(* IEC 61131-3 sources: daoli-st-library/DL_Motion (part 14) *)

(* ---- FB_DL_GearDecouple.st ---- *)
(*==============================================================================
 * 组件名称 (Component)  : FB_DL_GearDecouple
 * 所属子库 (Sublibrary) : DL_Motion
 * 当前版本 (Version)    : 1.0.0
 * 兼容性   (Platform)   : CODESYS 3.5+ / TwinCAT 3 / 汇川 InoProShop / 施耐德 Machine Expert
 *                         仅依赖 Standard.library（ABS），零厂商私有库
 * 功能描述 (Function)   : 电子齿轮渐变脱耦（MC_GearOut 语义）：耦合期输出比例
 *                         fRatioOut = iNum ÷ iDen；脱耦请求（bCoupled 下降沿）
 *                         后比例按 tRamp 渐降至 1:1（禁直接跳断，规格指定），
 *                         到达 1:1 置 bReleased（电平指示，重耦合撤销）；脱耦
 *                         斜坡中重新耦合（bCoupled 上升沿）比例斜坡回升至全
 *                         比例，无阶跃。iDen = 0 → 拒绝并锁存故障（除数前置
 *                         闸，规格指定）。
 * 接口     (Interface)  : 输入 bCoupled 耦合命令（TRUE=全比例耦合）、iNum 齿轮
 *                         分子、iDen 齿轮分母（域 <> 0）、fRampS 脱耦渐变时长
 *                         （域 > 0） [s]、fCycle 扫描周期（<=0 用缺省） [s]、
 *                         bReset 复位；输出 fRatioOut 渐变比例、bReleased
 *                         脱耦完成指示（电平）、bRamping 斜坡执行中指示、
 *                         eErrCode 错误码、bError 故障标志。
 * 边界     (Boundary)   : ① **属主边界（写死）：本件只出渐变比例标量，不接管
 *                         轴使能、不下齿轮指令**；齿轮耦合执行归
 *                         `FB_DL_ElectronicGear`。
 *                         ② 斜率口径：全比例 fRatioFull = iNum/iDen，斜坡速率
 *                         = (fRatioFull − 1) ÷ fRampS [1/s]；单步 = 速率 × fCy，
 *                         步内可达即贴目标（无过冲）；fRampS 用 LREAL 秒口径，
 *                         避免跨平台 TIME→实数转换链（R64 交付门槛规避，头注释
 *                         声明工程取舍）。
 *                         ③ fRatioFull = 1（1:1 齿轮）时斜坡速率恒 0：脱耦
 *                         请求即达 1:1，当拍 bReleased（无跳变路径，比例本就
 *                         不变）。
 *                         ④ 斜坡中禁直接跳断：bCoupled 变化只改目标值，输出
 *                         恒限步逼近（头注释声明，规格指定）。
 *                         ⑤ 组态闸：iDen = 0 或 fRampS <= 0 → 锁存故障，输出
 *                         冻结保持末值（比例冻结语义声明：R191 二选一之「冻结
 *                         保持」，故障期禁跳变），解除沿 = bReset 上升沿。
 *                         ⑥ 非有限判据（R79 双判）：fCycle 非有限按缺省周期
 *                         处理并入组态闸（iNum/iDen 整型无浮点域）。
 *                         ⑦ 零全局耦合（无 GVL / VAR_EXTERNAL / 物理地址）。
 * 分工声明 (Scope)      : 与 `FB_DL_ElectronicGear` 分工：恒比例齿轮耦合归那件、
 *                         渐变脱耦编排归本件；与 `FB_DL_AxisSynchronizedStop`
 *                         分工：同步停止归那件。
 * 来源标签 (Source Tag) : T1-6 ◐（PLCopen MC 语义只借 GearOut 脱耦完成语义，
 *                         斜坡渐变实现为道莅自研 clean-room）
 * 码表     (Codes)      : 本件不占用任何全局数字码位。出口为 LREAL 比例 +
 *                         BOOL 组 + ENUM 错误码；数字码位待主控收口阶段统一
 *                         派号。
 * 红线自检 (Redline)    : R1 ✓ 零 GVL/VAR_EXTERNAL ｜ R2 ✓ 零 %I/%Q/%M ｜ R3 ✓ 纯 IEC 61131-3
 *                         R4 ✓ 除数前置闸 + 限步逼近 + 故障冻结声明 ｜ R5 ✓ 声明逐行同行双语注释
 *                         R6 N/A（锁存态无 CASE 状态机） ｜ R7 ✓ 一 R_TRIG 段 0 无条件刷新
 * 修订历史 (Revision)   : 2026-11-20  v1.0.0  R50 首版（批次 3 · 序号 14）
 * 验收向量 (Acceptance) : ① iNum=2, iDen=1（全比例 2.0），fRampS=2.0，
 *                         fCycle=0.01 → 单步 0.005：脱耦后 200 拍达 1.0 →
 *                         bReleased=TRUE；② 100 拍时重耦合 → 比例自 1.5 反向
 *                         斜坡回升至 2.0（无阶跃）；③ iDen=0 → 锁存 eCfgBad，
 *                         fRatioOut 冻结末值；④ iNum=1, iDen=1 → 脱耦请求
 *                         当拍 fRatioOut=1.0、bReleased=TRUE。
 *==============================================================================*)

(*-----------------------------------------------------------------------------
 * 枚举: E_DL_GdcErr（错误码；故障级恒伴 bError=TRUE）
 *----------------------------------------------------------------------------*)
TYPE E_DL_GdcErr :
(
    eOk     := 0,   // 正常 / Normal
    eCfgBad := 1    // 故障级：分母零或斜坡时长非法（输出冻结保持） / Fault: zero denominator or bad ramp time
);
END_TYPE

FUNCTION_BLOCK FB_DL_GearDecouple
VAR_INPUT
    bCoupled : BOOL := TRUE;          // 耦合命令（TRUE=全比例，FALSE=脱耦请求） [-] / Coupled command
    iNum     : DINT := 2;             // 齿轮分子 [-] / Gear numerator
    iDen     : DINT := 1;             // 齿轮分母，域 <> 0 [-] / Gear denominator, must not be zero
    fRampS   : LREAL := 2.0;          // 脱耦渐变时长（全比例→1:1），域 > 0 [s] / Decouple ramp duration [s]
    fCycle   : LREAL := 0.0;          // 扫描周期（<=0 用缺省） [s] / Scan cycle, default used when <= 0
    bReset   : BOOL := FALSE;         // 复位，上升沿清组态锁存并回全比例/1:1 目标重算 [-] / Reset, rising edge clears latch
END_VAR
VAR_OUTPUT
    fRatioOut : LREAL;                // 渐变比例输出（限步逼近目标） [-] / Ramped ratio output
    bReleased : BOOL;                 // 脱耦完成指示（比例达 1:1 ∧ 脱耦请求中，电平） [-] / Released indicator, level
    bRamping  : BOOL;                 // 斜坡执行中指示 [-] / Ramping indicator
    eErrCode  : E_DL_GdcErr;          // 错误码出口 / Error code outlet
    bError    : BOOL;                 // 故障标志（组态锁存） [-] / Error flag, latched
END_VAR
VAR
    _fRatio   : LREAL := 1.0;         // 比例内部锁存（限步源，初值 1:1 安全态） / Ratio internal latch
    _fFull    : LREAL;                // 全比例 = iNum ÷ iDen（分母已闸） [-] / Full ratio
    _fRate    : LREAL;                // 斜坡速率（全比例−1）÷fRampS [1/s] / Ramp rate
    _fStep    : LREAL;                // 当拍最大步长 [1/拍] / Max step this scan
    _fTarget  : LREAL;                // 当拍目标比例 [-] / Target ratio this scan
    _fCy      : LREAL;                // 当拍有效周期 [s] / Effective cycle this scan
    _bCfgBad  : BOOL;                 // 组态非法当拍量 [-] / Illegal configuration
    _bErrLatch: BOOL;                 // 组态故障锁存位（解除沿 = bReset 上升沿） / Latched config fault
    rtReset   : R_TRIG;               // 复位沿实例，段 0 无条件调用 / Reset edge instance
END_VAR
VAR CONSTANT
    DL_GDC_CYDEF : LREAL := 0.01;     // 缺省扫描周期 [s] / Default scan cycle
    DL_GDC_ONE   : LREAL := 1.0;      // 1:1 基准与到达容差中心 [-] / Unity ratio base
    DL_GDC_ZERO  : LREAL := 0.0;      // 判零基准 [-] / Zero base
    DL_GDC_TOL   : LREAL := 1.0E-6;   // 到达判据容差（浮点禁 = 判等） [-] / Arrival tolerance
END_VAR

(* —— 段 0：非有限判 + 组态闸 + 周期派生 + 沿刷新 —— *)
IF fCycle <> fCycle THEN
    _fCy := DL_GDC_CYDEF;                          // 周期非有限按缺省（规格⑥） / Non-finite cycle to default
ELSIF fCycle > DL_GDC_ZERO THEN
    _fCy := fCycle;                                // 组态周期有效 / Configured cycle
ELSE
    _fCy := DL_GDC_CYDEF;                          // 周期缺省兜底 / Default fallback
END_IF
_bCfgBad := (iDen = 0) OR (fRampS <= DL_GDC_ZERO);   // 组态域闸（除数前置 + 斜坡时长） / Configuration gate
rtReset(CLK := bReset);                            // 复位沿，每拍必调 / Reset edge, every scan

(* —— 段 1：复位沿与组态锁存 —— *)
IF rtReset.Q THEN
    _bErrLatch := FALSE;                           // 清组态锁存（R188 声明：解除沿 = bReset 上升沿） / Clear cfg latch
END_IF
IF _bCfgBad AND (NOT _bErrLatch) THEN
    _bErrLatch := TRUE;                            // 锁存 / Latch
END_IF

(* —— 段 2：目标与速率派生（故障期跳过派生，冻结保持） —— *)
IF NOT _bErrLatch THEN
    _fFull := DINT_TO_LREAL(iNum) / DINT_TO_LREAL(iDen);   // 全比例（分母已闸，无除零） / Full ratio
    _fRate := ABS(_fFull - DL_GDC_ONE) / fRampS;   // 斜坡速率（对称双向同一速率） / Ramp rate
    _fStep := _fRate * _fCy;                       // 单步上限 [1/拍] / Max step
    IF bCoupled THEN
        _fTarget := _fFull;                        // 耦合目标 = 全比例 / Coupled target
    ELSE
        _fTarget := DL_GDC_ONE;                    // 脱耦目标 = 1:1（MC_GearOut 语义） / Decouple target
    END_IF
END_IF

(* —— 段 3：限步逼近（斜坡中禁直接跳断，规格④；步内可达即贴目标） —— *)
IF NOT _bErrLatch THEN
    IF _fTarget > (_fRatio + _fStep) THEN
        _fRatio := _fRatio + _fStep;               // 正向限步（重耦合回升无阶跃） / Ramp up limited
    ELSIF _fTarget < (_fRatio - _fStep) THEN
        _fRatio := _fRatio - _fStep;               // 负向限步（脱耦渐降） / Ramp down limited
    ELSE
        _fRatio := _fTarget;                       // 步内到达：贴目标 / Settle at target
    END_IF
END_IF

(* —— 段 4：出口单点映射（名实双出口同源，R191） —— *)
fRatioOut := _fRatio;                              // 比例出口（故障期冻结保持末值，头注释⑤声明） / Ratio outlet, frozen on fault
IF (NOT _bErrLatch) AND (NOT bCoupled)
   AND (ABS(_fRatio - DL_GDC_ONE) < DL_GDC_TOL) THEN
    bReleased := TRUE;                             // 脱耦完成电平（比例达 1:1 ∧ 脱耦请求中） / Released level
ELSE
    bReleased := FALSE;                            // 未完成/重耦合/故障期撤销 / Not released
END_IF
bRamping := (NOT _bErrLatch)
        AND (ABS(_fRatio - _fTarget) >= DL_GDC_TOL);   // 斜坡执行中（与目标距离超容差） / Ramping indicator
IF _bErrLatch THEN
    bError := TRUE;                                // 故障标志（R45 配对） / Error flag
    eErrCode := E_DL_GdcErr.eCfgBad;               // 故障级码 / Fault code
ELSE
    bError := FALSE;                               // 无故障级条件 / No fault
    eErrCode := E_DL_GdcErr.eOk;                   // 正常码 / OK code
END_IF

END_FUNCTION_BLOCK

(* ---- FB_DL_GearHobAxialShiftSeq.st ---- *)
//==============================================================================
// 功能块：FB_DL_GearHobAxialShiftSeq ｜ 中文名称：滚齿机滚刀轴向窜刀顺控（复杂度 C4）
// 所属子库：DL_Motion ｜ 版本 VERSION: v1.0.0 ｜ 兼容：CODESYS V3.5+ / TwinCAT 3 / 汇川 InoProShop
// 功能描述：滚刀磨损后沿刀轴窜动一个切削区宽度换新切削区——松刀轴夹紧 → 轴向进给
//           到目标位 → 到位稳定 → 重新夹紧确认 → 对刀校验 → 完成，累计窜刀量在完成
//           拍提交；超可用行程拒动、未松夹不得进给、未夹紧不得对刀、步超时落故障；
//           中止走两段化（先停进给 → 轴静止窗 → 再按安全序重新夹紧）。
// 开源溯源 (Origin)：道莅原创实现（参考 GB/T 1356 圆柱齿轮滚齿工艺与滚刀轴向窜刀
//           量工程惯例 分类与参数域，许可证=MIT，借鉴点=「按切削区宽度分步窜刀并
//           累计至刀轴可用行程上限」的工艺序）
// 单位表：长度[mm] / 时间[ms] / 计数[次]
// 错误码表（Motion 段 0008，故障窗口 0A01~0A08，信息窗口 0101）：
//   16#0008_0A01 故障级：组态非法（步长/上限/容差 <= 0、累计初值 < 0、时间量 <= 0）
//   16#0008_0A02 故障级：目标位 > fMaxTravelMm，拒动并置 xTravelLimit
//   16#0008_0A03 故障级：松夹相超时未到位，或进给期松夹信号丢失，禁进给
//   16#0008_0A04 故障级：夹紧相或中止再夹紧窗超时未确认，禁对刀
//   16#0008_0A05 故障级：进给步超时，或稳定窗满仍未判轴到位
//   16#0008_0A06 故障级：轴位置入口非有限（NaN / Inf）或幅值超合法上限，拒算
//   16#0008_0A07 故障级：对刀校验偏差 > fPosTolMm
//   16#0008_0A08 故障级兜底：状态机落 ELSE 非法态，全输出断
//   16#0008_0101 信息级：单步窜刀完成（完成拍，不置 bError）
//           故障级码全部锁存回放（R187），唯一清除路径 = bReset 上升沿。
// 状态机：E_DL_HobShiftState（八态：eIdle=0 / eRelease=10 / eShift=20 / eSettle=30 /
//           eReclamp=40 / eVerify=50 / eDone=60 / eFault=99）。八态为纯相序机，中止
//           两段化不占相位（八态契约锁定），由内部段号 _uAbortStage 驱动（0 无 /
//           1 已停进给待轴静止 / 2 再夹紧中）。
// 边界行为：① 组态非法与入口非有限一律锁存故障，故障相不按当下输入重推断；② 故障
//           相迁出唯一路径 = bReset 上升沿且组态合法、未超程；③ 中止段 A 拍内
//           xCmdMove 立即断、夹紧两命令均不动（O 型中位液压锁保持），机检断言：中止
//           段 A 不得出现 xClampCmd / xUnclampCmd 置位；④ 八态 CASE 每态显式 + ELSE
//           兜底 → 0A08 全断；⑤ 目标位在启动拍锁定一次。
// 语义假设：① fTotalShiftMm 为累计窜刀量初值，只在首扫且未窜过刀时载入内部累计量，
//           运行期不参与运算（避免累计量双属主），掉电保持由上层把 fShiftUsedMm 回写
//           该引脚，且只允许在 eIdle 且 xStart = FALSE 期间回写；② 夹紧电磁阀为双电控
//           O 型中位机能——两命令全 FALSE 时液压锁保持，故故障相「全输出断」不会松开
//           刀轴；③ 位置反馈为刀轴轴向绝对位 [mm]，正方向为离开主轴端面的窜刀方向。
// 依赖纪律：仅 Standard.library（TON / R_TRIG）；零 GVL、零 VAR_EXTERNAL、零物理地
//           址直连，业务侧只经引脚注入。
// 修订历史：v1.0.0 2026-11-25 R88 首版（无人值守批次 · 复杂件 C4 · 序号 1）
//==============================================================================

(*------------------------------------------------------------------------------
 * 枚举: E_DL_HobShiftState（归属本功能块，同文件发布，全库唯一定义）
 * 含义: 窜刀顺控相位，与段 8 输出置位、段 9 码映射一一对应。
 *-----------------------------------------------------------------------------*)
TYPE E_DL_HobShiftState :
(
    eIdle    := 0,   // 空闲：等启动沿 / Idle, awaiting the start edge
    eRelease := 10,  // 松夹：发松开命令并等松开到位 / Release the arbor clamp and wait for feedback
    eShift   := 20,  // 轴向进给：发运动命令至目标位 / Axial feed towards the target position
    eSettle  := 30,  // 到位稳定：等稳定窗与到位标志 / Settle, stability window and in-position flag
    eReclamp := 40,  // 夹紧确认：发夹紧命令并等夹紧反馈 / Reclamp and wait for clamp feedback
    eVerify  := 50,  // 对刀校验：实测位与目标位比对 / Tool-position verification against the target
    eDone    := 60,  // 完成：累计窜刀量已提交 / Done, accumulated shift committed
    eFault   := 99   // 故障：组态/超程/联锁/超时/非法态 / Fault, configuration, travel, interlock, timeout or illegal state
);
END_TYPE

FUNCTION_BLOCK FB_DL_GearHobAxialShiftSeq
VAR_INPUT
    xEnable       : BOOL;   // 使能，FALSE 期间按中止处理 [—] / Enable, a drop is treated as an abort
    xStart        : BOOL;   // 启动请求，上升沿生效 [—] / Start request, rising edge effective
    xAbort        : BOOL;   // 中止请求，任意拍生效 [—] / Abort request, effective on any scan
    xReset        : BOOL;   // 故障复位，上升沿清全部锁存 [—] / Fault reset, rising edge clears all latches
    fShiftStepMm  : LREAL;  // 单步窜刀量 [mm]，须 > 0 / Per-step axial shift [mm], must be > 0
    fTotalShiftMm : LREAL;  // 累计窜刀量初值 [mm]，仅首扫载入 / Initial accumulated shift [mm], first scan only
    fAxisPosMm    : LREAL;  // 刀轴实际轴向位置 [mm] / Hob arbor actual axial position [mm]
    xAxisInPos    : BOOL;   // 轴到位标志 [—] / Axis in-position flag
    xClampClosed  : BOOL;   // 夹紧到位反馈 [—] / Clamp-closed feedback
    xClampOpen    : BOOL;   // 松开到位反馈 [—] / Clamp-open feedback
    tMoveTimeout  : TIME;   // 进给/校验步超时 [ms] / Feed and verification step timeout [ms]
    tSettleTime   : TIME;   // 到位稳定窗 [ms] / In-position settle window [ms]
    fPosTolMm     : LREAL;  // 对刀位置容差 [mm]，须 > 0 / Verification position tolerance [mm]
    fMaxTravelMm  : LREAL;  // 刀轴可用窜刀总行程 [mm] / Total usable axial shift travel [mm]
END_VAR
VAR_OUTPUT
    xCmdMove      : BOOL;   // 轴向进给命令 [—] / Axial feed command
    fCmdPosMm     : LREAL;  // 目标位命令 [mm] / Target position command [mm]
    xClampCmd     : BOOL;   // 夹紧命令（双电控 O 型中位，断电保持） [—] / Clamp command, O-centre holds on power loss
    xUnclampCmd   : BOOL;   // 松开命令（双电控 O 型中位，断电保持） [—] / Unclamp command, holds on power loss
    bRunning      : BOOL;   // 顺控运行中（非空闲非完成非故障非中止） [—] / Sequencing active
    bDone         : BOOL;   // 单步窜刀完成相电平 [—] / Single shift step done, level in the done phase
    bError        : BOOL;   // 故障级标志，仅故障级码置位 [—] / Fault-class flag, fault-level codes only
    nErrCode      : UDINT;  // 错误码，0 = 无错 [—] / Error code, 0 = none
    fShiftUsedMm  : LREAL;  // 累计窜刀量出口 [mm] / Accumulated axial shift outlet [mm]
    nShiftCount   : UDINT;  // 累计窜刀次数 [次] / Accumulated shift step count
    xTravelLimit  : BOOL;   // 窜刀行程上限已达（拒动锁存） [—] / Travel limit reached, refuse-to-move latch
END_VAR
VAR
    _eState       : E_DL_HobShiftState := E_DL_HobShiftState.eIdle; // 当前相位 [—] / Current phase
    _bInit        : BOOL := FALSE;      // 首扫标志，取非判定 [—] / First-scan flag, tested negated
    _fShiftUsedMm : LREAL;              // 内部累计窜刀量 [mm] / Internal accumulated shift [mm]
    _fTargetPosMm : LREAL;              // 本步目标位 [mm] = 累计 + 步长 / Step target [mm] = accumulated + step
    _fPosPrevMm   : LREAL;              // 上拍轴位快照 [mm]，静止判据用 / Previous-scan position [mm]
    _nShiftCount  : UDINT;              // 内部累计窜刀次数 [次] / Internal shift step counter
    _bCfgBad      : BOOL;               // 组态非法锁存 / Illegal configuration latch
    _bCfgOk       : BOOL;               // 本拍组态合法（派生量不锁存） [—] / Configuration legal this scan, derived
    _bAxisBad     : BOOL;               // 轴位置非有限锁存 / Non-finite axis position latch
    _bOverTravel  : BOOL;               // 超窜刀行程锁存 / Over-travel latch
    _bReleaseTmo  : BOOL;               // 松夹未到位/信号丢失锁存 / Release-not-reached latch
    _bClampTmo    : BOOL;               // 夹紧未确认锁存 / Clamp-not-confirmed latch
    _bFeedTmo     : BOOL;               // 进给步超时锁存 / Feed step timeout latch
    _bVerifyErr   : BOOL;               // 对刀超差锁存 / Verification error latch
    _bIllegal     : BOOL;               // 非法状态标志 / Illegal state flag
    _bInfoDone    : BOOL;               // 单步完成信息当拍标志 / Step-done info flag of this scan
    _bAbortReq    : BOOL;               // 中止请求合成（xAbort 或失能） [—] / Combined abort request
    _bFeedPermit  : BOOL;               // 进给许可（松开到位且未夹紧） [—] / Feed permit, released and not clamped
    _bStandstill  : BOOL;               // 轴静止判据（本拍位移小于阈值） [—] / Axis standstill criterion
    _uAbortStage  : UINT;               // 中止段号 0=无 1=待静止 2=再夹紧 / Abort stage 0 none 1 standstill 2 reclamp
    rtStart       : R_TRIG;             // 启动沿，段 5 无条件刷新 [—] / Start edge, refreshed in segment 5
    rtReset       : R_TRIG;             // 复位沿，段 5 无条件刷新 [—] / Reset edge, refreshed in segment 5
    tonRelease    : TON;                // 松夹相超时计时 [ms] / Release phase timeout [ms]
    tonMove       : TON;                // 进给相超时计时 [ms] / Feed phase timeout [ms]
    tonSettle     : TON;                // 稳定窗计时 [ms] / Settle window timer [ms]
    tonReclamp    : TON;                // 夹紧确认超时计时 [ms] / Reclamp timeout [ms]
    tonVerify     : TON;                // 对刀校验超时计时 [ms] / Verification timeout [ms]
    tonStandstill : TON;                // 中止段 A 静止窗计时 [ms] / Abort stage A standstill window [ms]
    tonAbortClamp : TON;                // 中止段 B 再夹紧确认窗计时 [ms] / Abort stage B reclamp window [ms]
END_VAR
VAR CONSTANT
    DL_EPS           : LREAL := 1.0E-9;      // 浮点容差零点，兼作除法分母下限 / Float epsilon, also the divisor floor
    DL_HOB_STILL_MM  : LREAL := 0.005;       // 静止窗每拍位移阈值 [mm] / Per-scan displacement threshold [mm]
    DL_HOB_ABORT_T   : TIME  := T#1500MS;    // 中止静止窗时长 [ms] / Abort standstill window [ms]
    DL_HOB_CLAMP_T   : TIME  := T#3000MS;    // 中止再夹紧确认窗 [ms] / Abort reclamp confirm window [ms]
    DL_HOB_POS_MAX   : LREAL := 1.0E9;       // 位置幅值合法上限 [mm] / Legal position magnitude ceiling [mm]
END_VAR

(*------------------------------------------------------------------------------
 * 段 1｜每拍预置：全部输出先落安全侧，单拍标志预清零
 *      All outputs preset to the safe side, one-shot flags pre-cleared
 *-----------------------------------------------------------------------------*)
xCmdMove := FALSE;  fCmdPosMm := 0.0;       // 进给命令与目标位先清 / Feed command and target cleared first
xClampCmd := FALSE; xUnclampCmd := FALSE;   // 夹紧两命令先断（O 型中位保持） / Both clamp commands cleared, O-centre holds
bRunning := FALSE;  bDone := FALSE;         // 运行与完成标志每拍重算 / Running and done flags recomputed
bError := FALSE;    nErrCode := 16#0000_0000; // 故障标志与错误码每拍重算 / Fault flag and code recomputed
xTravelLimit := FALSE;                      // 超程标志每拍重算 / Travel limit flag recomputed
_bIllegal := FALSE; _bInfoDone := FALSE;    // 非法态与完成信息预清零 / Illegal and done-info flags pre-cleared

(*------------------------------------------------------------------------------
 * 段 2｜首扫初始化：相位、累计量、计数与中止段号复位
 *      First-scan initialisation of phase, accumulated shift, counter and abort stage
 *-----------------------------------------------------------------------------*)
IF NOT _bInit THEN
    _eState       := E_DL_HobShiftState.eIdle;   // 相位从空闲起步 / Phase starts idle
    _fShiftUsedMm := 0.0;  _fTargetPosMm := 0.0; // 累计量与目标位先清零 / Accumulated shift and target at zero
    _fPosPrevMm   := 0.0;  _nShiftCount  := 0;   // 位置快照与窜刀计数清零 / Position snapshot and counter at zero
    _uAbortStage  := 0;                          // 中止段号从零起步 / Abort stage starts at zero
    _bInit        := TRUE;                       // 首扫只做一次 / The first scan runs once
END_IF

(*------------------------------------------------------------------------------
 * 段 3｜入口非有限闸 + 组态闸 + 目标位预计算 + 超行程拒动判定
 *      Non-finite inlet gate, configuration gates, target computation, travel check
 *-----------------------------------------------------------------------------*)
IF NOT (fAxisPosMm > -1.0E30 AND fAxisPosMm < 1.0E30) THEN _bAxisBad := TRUE; END_IF    // 轴位非有限 → 0A06 / Non-finite position, 0A06
IF ABS(fAxisPosMm) > DL_HOB_POS_MAX THEN _bAxisBad := TRUE; END_IF                     // 轴位幅值超上限 → 0A06 / Beyond the ceiling, 0A06
IF NOT (fShiftStepMm > -1.0E30 AND fShiftStepMm < 1.0E30) THEN _bCfgBad := TRUE; END_IF  // 步长非有限 → 0A01 / Non-finite step, 0A01
IF NOT (fMaxTravelMm > -1.0E30 AND fMaxTravelMm < 1.0E30) THEN _bCfgBad := TRUE; END_IF // 行程上限非有限 → 0A01 / Non-finite limit, 0A01
IF NOT (fPosTolMm > -1.0E30 AND fPosTolMm < 1.0E30) THEN _bCfgBad := TRUE; END_IF      // 容差非有限 → 0A01 / Non-finite tolerance, 0A01
IF NOT (fTotalShiftMm > -1.0E30 AND fTotalShiftMm < 1.0E30) THEN _bCfgBad := TRUE; END_IF // 累计初值非有限 → 0A01 / Non-finite initial shift, 0A01
IF (fShiftStepMm <= DL_EPS) OR (fMaxTravelMm <= DL_EPS) OR (fPosTolMm <= DL_EPS) THEN _bCfgBad := TRUE; END_IF // 三者须为正 → 0A01 / All three must be positive
IF fTotalShiftMm < 0.0 THEN _bCfgBad := TRUE; END_IF                                   // 累计初值负值非法 → 0A01 / Negative initial shift, 0A01
IF (tMoveTimeout <= T#0MS) OR (tSettleTime <= T#0MS) THEN _bCfgBad := TRUE; END_IF      // 时间量须为正 → 0A01 / Time values must be positive
_bCfgOk := NOT _bCfgBad;                    // 本拍组态合法派生量 / Configuration-legal derived flag of this scan
IF (_nShiftCount = 0) AND (_eState = E_DL_HobShiftState.eIdle) AND (NOT _bCfgBad) THEN
    _fShiftUsedMm := fTotalShiftMm;         // 累计初值载入（仅未窜过刀时） / Initial shift loaded before the first step
END_IF
IF (_eState = E_DL_HobShiftState.eIdle) OR (_eState = E_DL_HobShiftState.eDone)
   OR (_eState = E_DL_HobShiftState.eFault) THEN
    _fTargetPosMm := _fShiftUsedMm + fShiftStepMm; // 目标位 = 累计窜刀量 + 步长 [mm]，仅非运行相更新，运行期锁定 / Target updated outside running phases only
END_IF
IF (_bCfgOk) AND (NOT _bAxisBad) AND (_fTargetPosMm > fMaxTravelMm) THEN
    _bOverTravel := TRUE;                   // 目标位超可利用行程，拒动锁存 → 0A02 / Beyond usable travel, 0A02
END_IF

(*------------------------------------------------------------------------------
 * 段 4｜中止入口（段 0→1）、静止判据与复位
 *      Abort entry, standstill criterion and the reset edge
 *-----------------------------------------------------------------------------*)
_bAbortReq   := xAbort OR (NOT xEnable);    // 中止请求合成：显式中止或失能 / Combined abort: explicit abort or enable loss
_bFeedPermit := xClampOpen AND (NOT xClampClosed); // 进给许可：松开到位且未夹紧 / Feed permit: released and not clamped
IF _bAbortReq AND (_uAbortStage = 0) AND (_eState <> E_DL_HobShiftState.eIdle)
   AND (_eState <> E_DL_HobShiftState.eDone) AND (_eState <> E_DL_HobShiftState.eFault) THEN
    _uAbortStage := 1;                      // 进中止段 A：先停进给待轴静止 / Enter abort stage A, await standstill
END_IF
_bStandstill := ABS(fAxisPosMm - _fPosPrevMm) < DL_HOB_STILL_MM; // 本拍位移小于阈值视为静止 / A per-scan move below the threshold is standstill
IF rtReset.Q THEN
    _bCfgBad := FALSE;  _bAxisBad := FALSE; _bOverTravel := FALSE; // 复位清组态/非有限/超程锁存 / Clears configuration, non-finite and travel
    _bReleaseTmo := FALSE; _bClampTmo := FALSE; _bFeedTmo := FALSE; // 复位清松夹/夹紧/超时锁存 / Clears release, clamp and timeout
    _bVerifyErr := FALSE;                   // 复位清对刀校验锁存 / Clears the verification latch
END_IF

(*------------------------------------------------------------------------------
 * 段 5｜定时器与边沿无条件周期刷新（R7：CASE 之外每拍必调，各司其职不复用）
 *      Timers and edges refreshed unconditionally every scan, outside the CASE
 *-----------------------------------------------------------------------------*)
rtStart(CLK := xStart);                     // 启动沿刷新 / Start edge refreshed
rtReset(CLK := xReset);                     // 复位沿刷新 / Reset edge refreshed
tonRelease(IN := (_eState = E_DL_HobShiftState.eRelease) AND (_uAbortStage = 0), PT := tMoveTimeout); // 松夹相超时 / Release timeout
tonMove(IN := (_eState = E_DL_HobShiftState.eShift) AND (_uAbortStage = 0), PT := tMoveTimeout);      // 进给相超时 / Feed timeout
tonSettle(IN := (_eState = E_DL_HobShiftState.eSettle) AND (_uAbortStage = 0), PT := tSettleTime);    // 稳定窗计时 / Settle window
tonReclamp(IN := (_eState = E_DL_HobShiftState.eReclamp) AND (_uAbortStage = 0), PT := tMoveTimeout); // 夹紧确认超时 / Reclamp timeout
tonVerify(IN := (_eState = E_DL_HobShiftState.eVerify) AND (_uAbortStage = 0), PT := tMoveTimeout);   // 对刀校验超时 / Verification timeout
tonStandstill(IN := (_uAbortStage = 1) AND _bStandstill, PT := DL_HOB_ABORT_T); // 中止段 A 静止窗 / Abort stage A standstill window
tonAbortClamp(IN := (_uAbortStage = 2), PT := DL_HOB_CLAMP_T);                  // 中止段 B 再夹紧窗 / Abort stage B reclamp window

(*------------------------------------------------------------------------------
 * 段 6｜中止段推进（1→2 轴静止后按安全序再夹紧，2→0 收口）
 *      Abort stage progression, reclamp only after the axis is standstill
 *-----------------------------------------------------------------------------*)
IF (_uAbortStage = 1) AND tonStandstill.Q THEN
    _uAbortStage := 2;                      // 轴静止窗满，进再夹紧段 / Standstill elapsed, enter reclamp
END_IF
IF _uAbortStage = 2 THEN
    IF xClampClosed THEN
        _uAbortStage := 0;                  // 再夹紧已确认，中止收口 / Reclamp confirmed, abort closed
        _eState      := E_DL_HobShiftState.eIdle; // 回空闲 / Back to idle
    ELSIF tonAbortClamp.Q THEN
        _bClampTmo   := TRUE;               // 再夹紧窗满无反馈 → 0A04 / Window elapsed without feedback, 0A04
        _uAbortStage := 0;                  // 中止段收口 / Abort stage closed
        _eState      := E_DL_HobShiftState.eFault; // 落故障 / Fall to fault
    END_IF
END_IF

(*------------------------------------------------------------------------------
 * 段 7｜状态机（中止期间迁移冻结；本段只做迁移，输出在段 8）
 *      Phase machine, transitions frozen while aborting, outputs in segment 8
 *-----------------------------------------------------------------------------*)
IF _uAbortStage = 0 THEN
    CASE _eState OF
        E_DL_HobShiftState.eIdle:           // 空闲：启动沿 + 组态合法 + 未超程才进松夹 / Idle, legal start edge only
            IF rtStart.Q AND _bCfgOk AND (NOT _bAxisBad) AND (NOT _bOverTravel) AND (NOT _bAbortReq) THEN
                _fTargetPosMm := _fShiftUsedMm + fShiftStepMm; // 启动拍锁定目标位 / Target locked at the start edge
                _eState := E_DL_HobShiftState.eRelease;        // 进松夹相 / To the release phase
            END_IF
        E_DL_HobShiftState.eRelease:        // 松夹：松开到位才允许进给 / Release, feeding only once released
            IF _bFeedPermit THEN _eState := E_DL_HobShiftState.eShift; // 松开到位，进进给相 / Released, to feed
            ELSIF tonRelease.Q THEN _bReleaseTmo := TRUE; _eState := E_DL_HobShiftState.eFault; // 超时未到位 → 0A03 / Timeout, 0A03
            END_IF
        E_DL_HobShiftState.eShift:          // 进给：松夹信号丢失即故障，到位进稳定相 / Feed, permit loss faults
            IF NOT _bFeedPermit THEN _bReleaseTmo := TRUE; _eState := E_DL_HobShiftState.eFault; // 松夹丢失 → 0A03 / Permit lost, 0A03
            ELSIF xAxisInPos THEN _eState := E_DL_HobShiftState.eSettle; // 到位，进稳定相 / In position, to settle
            ELSIF tonMove.Q THEN _bFeedTmo := TRUE; _eState := E_DL_HobShiftState.eFault; // 进给步超时 → 0A05 / Feed timeout, 0A05
            END_IF
        E_DL_HobShiftState.eSettle:         // 稳定：稳定窗满且仍到位才进夹紧 / Settle, reclamp after the window
            IF tonSettle.Q AND xAxisInPos THEN _eState := E_DL_HobShiftState.eReclamp; // 稳定到位，进夹紧 / Stable, to reclamp
            ELSIF tonSettle.Q THEN _bFeedTmo := TRUE; _eState := E_DL_HobShiftState.eFault; // 窗满未到位 → 0A05 / Elapsed, 0A05
            END_IF
        E_DL_HobShiftState.eReclamp:        // 夹紧：夹紧确认才允许对刀校验 / Reclamp, verification only once clamped
            IF xClampClosed AND (NOT xClampOpen) THEN _eState := E_DL_HobShiftState.eVerify; // 夹紧确认，进校验 / Clamped, verify
            ELSIF tonReclamp.Q THEN _bClampTmo := TRUE; _eState := E_DL_HobShiftState.eFault; // 超时未夹紧 → 0A04 / Clamp timeout, 0A04
            END_IF
        E_DL_HobShiftState.eVerify:         // 对刀校验：夹紧须保持，偏差在容差内即完成 / Verify with the clamp held
            IF NOT xClampClosed THEN _bClampTmo := TRUE; _eState := E_DL_HobShiftState.eFault; // 夹紧丢失 → 0A04 / Clamp lost, 0A04
            ELSIF ABS(fAxisPosMm - _fTargetPosMm) <= fPosTolMm THEN
                _fShiftUsedMm := _fShiftUsedMm + fShiftStepMm; // 完成拍提交累计窜刀量 / Accumulated shift committed
                _nShiftCount := _nShiftCount + 1; _bInfoDone := TRUE; // 次数递增 + 完成信息 / Counter plus done info
                _eState := E_DL_HobShiftState.eDone;           // 进完成相 / To the done phase
            ELSIF tonVerify.Q THEN _bVerifyErr := TRUE; _eState := E_DL_HobShiftState.eFault; // 超差 → 0A07 / Deviation, 0A07
            END_IF
        E_DL_HobShiftState.eDone:           // 完成：启动撤销且无中止请求才回空闲 / Done, back to idle once start drops
            IF (NOT xStart) AND (NOT _bAbortReq) THEN _eState := E_DL_HobShiftState.eIdle; END_IF
        E_DL_HobShiftState.eFault:          // 故障：复位沿且组态合法且未超程才回空闲 / Fault, reset edge only
            IF rtReset.Q AND _bCfgOk AND (NOT _bAxisBad) AND (NOT _bOverTravel) THEN _eState := E_DL_HobShiftState.eIdle; END_IF
        ELSE                                // 非法状态兜底（R6：CASE 必带 ELSE）/ Illegal-state fallback
            _bIllegal := TRUE; _eState := E_DL_HobShiftState.eFault; // 非法态 → 0A08，落故障 / Illegal state, 0A08
    END_CASE
END_IF

(*------------------------------------------------------------------------------
 * 段 8｜输出置位（次序即安全：进给受许可闸，夹紧两命令互斥）
 *      Output assignment, feed gated by the permit, clamp commands exclusive
 *-----------------------------------------------------------------------------*)
CASE _eState OF
    E_DL_HobShiftState.eRelease:            // 松夹相：只发松开命令 / Release phase, unclamp only
        xUnclampCmd := TRUE;                // 松开命令 / Unclamp command
    E_DL_HobShiftState.eShift:              // 进给相：命令位 + 进给许可双重闸 / Feed phase, target plus permit
        fCmdPosMm := _fTargetPosMm;         // 目标位命令 / Target position command
        xCmdMove  := _bFeedPermit;          // 未松夹到位不得进给 / Feeding forbidden unless released
    E_DL_HobShiftState.eSettle:             // 稳定相：保持命令位不撤 / Settle phase, command held
        fCmdPosMm := _fTargetPosMm;         // 目标位保持 / Target position held
    E_DL_HobShiftState.eReclamp:            // 夹紧相：只发夹紧命令 / Reclamp phase, clamp only
        xClampCmd := TRUE;                  // 夹紧命令 / Clamp command
    E_DL_HobShiftState.eDone:               // 完成相：完成电平 / Done phase, done level
        bDone := TRUE;                      // 单步完成 / Single step done
    ELSE                                    // 其余相（空闲/校验/故障）全断 / Other phases, all off
        xCmdMove := FALSE; xClampCmd := FALSE; xUnclampCmd := FALSE; // 全输出断 / All outputs off
END_CASE
IF _uAbortStage >= 1 THEN
    xCmdMove    := FALSE;                   // 中止段 A：进给立即断（安全侧） / Abort A, feed cut immediately
    xClampCmd   := FALSE; xUnclampCmd := FALSE; // 静止窗内两夹紧命令均不动（O 型中位保持） / Both idle in the window
    fCmdPosMm   := _fTargetPosMm;           // 命令位保持，禁回零溜刀 / Command held, no return-to-zero creep
    IF _uAbortStage = 2 THEN
        xClampCmd := NOT xClampClosed;      // 中止段 B：未夹紧则发夹紧（安全序） / Abort B, clamp unless clamped
    END_IF
END_IF
bRunning := (_eState <> E_DL_HobShiftState.eIdle) AND (_eState <> E_DL_HobShiftState.eDone)
            AND (_eState <> E_DL_HobShiftState.eFault) AND (_uAbortStage = 0); // 运行标志 / Running flag

(*------------------------------------------------------------------------------
 * 段 9｜出口量与错误码映射（锁存回放，R187：故障相不按当下输入重推断）
 *      Outlet quantities and the error-code map, latched replay
 *-----------------------------------------------------------------------------*)
fShiftUsedMm := _fShiftUsedMm;              // 累计窜刀量出口 [mm] / Accumulated shift outlet [mm]
nShiftCount  := _nShiftCount;               // 窜刀次数出口 [次] / Shift count outlet
xTravelLimit := _bOverTravel;               // 超程拒动出口 / Travel-limit outlet
IF _bIllegal THEN nErrCode := 16#0008_0A08; bError := TRUE;        // 故障级兜底：非法态 / Fault, illegal state fallback
ELSIF _bCfgBad THEN nErrCode := 16#0008_0A01; bError := TRUE;      // 故障级：组态非法 / Fault, illegal configuration
ELSIF _bAxisBad THEN nErrCode := 16#0008_0A06; bError := TRUE;     // 故障级：轴位非有限 / Fault, non-finite position
ELSIF _bOverTravel THEN nErrCode := 16#0008_0A02; bError := TRUE;  // 故障级：超窜刀行程 / Fault, over travel
ELSIF _bReleaseTmo THEN nErrCode := 16#0008_0A03; bError := TRUE;  // 故障级：松夹不到位 / Fault, release not reached
ELSIF _bClampTmo THEN nErrCode := 16#0008_0A04; bError := TRUE;    // 故障级：夹紧未确认 / Fault, clamp not confirmed
ELSIF _bFeedTmo THEN nErrCode := 16#0008_0A05; bError := TRUE;     // 故障级：进给步超时 / Fault, feed step timeout
ELSIF _bVerifyErr THEN nErrCode := 16#0008_0A07; bError := TRUE;   // 故障级：对刀超差 / Fault, verification out of tolerance
ELSIF _bInfoDone THEN nErrCode := 16#0008_0101;                    // 信息级：单步完成，不置 bError / Info, step done
END_IF
_fPosPrevMm := fAxisPosMm;                  // 位置快照推进（供下拍静止判据） / Position snapshot advanced for the next scan
END_FUNCTION_BLOCK

(* ---- FB_DL_GearInPhaseAlign.st ---- *)
(*
  FB_DL_GearInPhaseAlign  —  电子齿轮啮合相位对齐（相位差窗 + 从轴偏置补偿） / Electronic gear-in phase alignment with phase-error window and slave offset compensation
  分类 Category : DL_Motion
  版本 Version  : 1.0.0
  来源 Source   : t1-6-plcopen — PLCopen Motion 接口映射层族深化
  溯源 Origin   : 道莅 clean-room 实现；从轴相位 = 主轴位置×传动比 + 偏置 为公开电子齿轮运动学关系，
                 本件仅做 MC_GearIn 前置相位判据与偏置补偿的映射层，不内联轨迹规划内核
  功能 Function : 1) 理想从轴相位 _fIdealDeg = fMasterPosDeg × fGearRatio；
                  2) 相位差 _fPhaseErrDeg = 归一化(fSlavePosDeg - _fIdealDeg - fPhaseTargetDeg)，
                  归一化按 ±360° 折算（除以常量 360.0，禁 MOD 非标准扩展）；
                  3) 判据：|相位差| <= fPhaseTolDeg → bInPhase（可啮合）；
                  4) 偏置补偿：补偿量按 -相位差 × fGainDegPerDeg 计算，钳制到
                  ±fOffsetMaxDeg 并限速（单次不超过 fOffsetStepDeg）；
                  5) 本件只有故障码、无信息码（派单硬约束）。
  接口 Interface: 输入主轴/从轴位置、传动比、目标相位、容差、偏置域；输出相位差与偏置
  边界 Boundary : ① 组态闸：fGearRatio <= 0.0、fPhaseTolDeg <= 0.0、fOffsetMaxDeg <= 0.0、
                  fOffsetStepDeg <= 0.0、fGainDegPerDeg <= 0.0 → 04A7 锁存；
                  ② 位置或传动比非有限（NaN 自反 + Inf 差值自减）→ 04A7 锁存，偏置冻结保持；
                  ③ 归一化除法除数为常量 360.0（无除零风险）；
                  ④ 一个 R_TRIG，段 0 无条件调用；⑤ 故障相迁出唯一路径 = bReset 上升沿；
                  ⑥ 零全局耦合：无 GVL / VAR_EXTERNAL / %I %Q %M 直接地址。
  依赖 Depends  : Standard.library（R_TRIG）
  码表 Error codes（Motion 段 0004，故障窗口 04A7；本件无信息码）:
    16#0004_04A7 故障级：相位对齐故障总码（组态非法 / 位置或传动比非有限），
                 锁存至 bReset 上升沿；归因见 eCause，不新增码位（派单硬约束单码）
  修订历史 Revision :
    2026-11-19  v1.0.0  R43 首版（批次 4 · 序号 19）
*)

TYPE E_DL_GpaState :
(
    eIdle   := 0,     // 未使能待对齐 / Idle, waiting alignment
    eAlign  := 10,    // 相位对齐中（偏置补偿） / Aligning with offset compensation
    eReady  := 20,    // 相位在窗：可啮合 / In phase, gear-in permitted
    eFault  := 90     // 故障锁存相（偏置冻结） / Fault latched, offset frozen
);
END_TYPE

TYPE E_DL_GpaCause :
(
    eNone       := 0, // 无故障成因 / No cause
    eCfgIllegal := 1, // 组态非法 / Illegal configuration
    eNonFinite  := 2  // 输入非有限 / Non-finite input
);
END_TYPE

FUNCTION_BLOCK FB_DL_GearInPhaseAlign
VAR_INPUT
    fMasterPosDeg  : REAL := 0.0;      // 主轴位置 [°] / Master position
    fSlavePosDeg   : REAL := 0.0;      // 从轴位置 [°] / Slave position
    fGearRatio     : REAL := 1.0;      // 传动比 [从轴°/主轴°]，域 > 0 / Gear ratio
    fPhaseTargetDeg: REAL := 0.0;      // 目标相位差 [°] / Target phase difference
    fPhaseTolDeg   : REAL := 2.0;      // 相位差窗 [°]，域 > 0 / Phase window
    fGainDegPerDeg : REAL := 0.8;      // 补偿增益 [°/°]，域 > 0 / Compensation gain
    fOffsetMaxDeg  : REAL := 30.0;     // 偏置限幅 [°]，域 > 0 / Offset limit
    fOffsetStepDeg : REAL := 5.0;      // 单周期偏置步长 [°]，域 > 0 / Offset step
    bEnable        : BOOL := FALSE;    // 对齐使能（电平）[-] / Alignment enable
    bReset         : BOOL := FALSE;    // 复位命令，上升沿清故障与偏置 [-] / Reset edge
END_VAR
VAR_OUTPUT
    eState         : E_DL_GpaState;    // 状态出口，段 6 单点映射 / State outlet
    eCause         : E_DL_GpaCause;    // 故障成因出口（R190） / Fault cause outlet
    fPhaseErrDeg   : REAL;             // 归一化相位差 [°] / Normalised phase error
    fOffsetDeg     : REAL;             // 从轴偏置补偿 [°] / Slave offset compensation
    bInPhase       : BOOL;             // 相位在窗（MC_GearIn 许可）[-] / In-phase permit
    bError         : BOOL;             // 故障锁存标志 [-] / Fault latch flag
    nErrId         : UDINT;            // 故障码，0 = 无故障（本件无信息码） / Fault code only
END_VAR
VAR
    _eState        : E_DL_GpaState := E_DL_GpaState.eIdle;   // 内部相位（CASE 唯一写入目标） / Internal phase
    _eCause        : E_DL_GpaCause := E_DL_GpaCause.eNone;   // 故障成因锁存（锁存量） / Latched cause
    rtReset        : R_TRIG;           // 复位沿实例，每周期无条件调用 / Reset edge
    _fOffsetDeg    : REAL;             // 偏置保持量（持久） / Offset holding slot
    _fIdealDeg     : REAL;             // 理想从轴相位 [°]（当拍量） / Ideal slave phase
    _fErrRawDeg    : REAL;             // 未归一化相位差 [°]（当拍量） / Raw phase error
    _fErrDeg       : REAL;             // 归一化相位差 [°]（当拍量） / Normalised phase error
    _fCmdDeg       : REAL;             // 目标偏置 [°]（当拍量） / Target offset
    _bInPhase      : BOOL;             // 相位在窗当拍量 [-] / In-phase verdict
    _bNonFin       : BOOL;             // 输入非有限当拍量 [-] / Non-finite input
    _bCfgBad       : BOOL;             // 组态非法当拍量 [-] / Config illegal
    _bFault        : BOOL;             // 故障锁存位（锁存量） / Latched fault bit
    _uFault        : UDINT;            // 故障码锁存（锁存量） / Latched fault code
END_VAR

(* —— 段 0：沿实例无条件周期刷新 + 相位差归一化（除数为常量 360.0） —— *)
_fIdealDeg := fMasterPosDeg * fGearRatio;                                    // 理想从轴相位 / Ideal slave phase
_fErrRawDeg := fSlavePosDeg - _fIdealDeg - fPhaseTargetDeg;                  // 未归一化相位差 / Raw phase error
_fErrDeg := _fErrRawDeg;                                                     // 归一化初值 / Normalisation start
IF _fErrDeg > 180.0 THEN                                                     // 超半周：折算到负半周 / Wrap to negative half
    _fErrDeg := _fErrDeg - 360.0;
ELSIF _fErrDeg < -180.0 THEN                                                 // 低于负半周：折算到正半周 / Wrap to positive half
    _fErrDeg := _fErrDeg + 360.0;
END_IF
_bInPhase := ABS(_fErrDeg) <= fPhaseTolDeg;                                  // 相位窗判据（容差式） / Phase window verdict
_bNonFin := (fMasterPosDeg <> fMasterPosDeg) OR (fSlavePosDeg <> fSlavePosDeg) OR (fGearRatio <> fGearRatio)
         OR ((fMasterPosDeg - fMasterPosDeg) <> (fMasterPosDeg - fMasterPosDeg))
         OR ((fSlavePosDeg - fSlavePosDeg) <> (fSlavePosDeg - fSlavePosDeg))
         OR ((fGearRatio - fGearRatio) <> (fGearRatio - fGearRatio));        // NaN 自反 + Inf 差值自减 / NaN and Inf
_bCfgBad := (fGearRatio <= 0.0) OR (fPhaseTolDeg <= 0.0) OR (fOffsetMaxDeg <= 0.0)
            OR (fOffsetStepDeg <= 0.0) OR (fGainDegPerDeg <= 0.0);           // 组态非法当拍量 / Config illegal
rtReset(CLK := bReset);                                                      // 复位沿，每拍必调 / Reset edge

(* —— 段 1：单拍量预清零（锁存量与偏置保持量不入清单） —— *)
fPhaseErrDeg := 0.0;               // 相位差出口缺省 0 / Phase error default
bInPhase := FALSE;                 // 在窗镜像缺省 FALSE（安全侧） / In-phase default safe
nErrId := 16#0000_0000;            // 故障码缺省无故障 / Fault code default

(* —— 段 2：复位沿 + 组态域闸 —— *)
IF rtReset.Q THEN                              // rtReset.Q = 当拍量 / current scan
    _bFault := FALSE;                          // 清故障锁存位（锁存量） / Clear fault latch
    _uFault := 16#0000_0000;                   // 清故障锁存码（锁存量） / Clear fault code
    _eCause := E_DL_GpaCause.eNone;            // 清成因（锁存量） / Clear cause
    _fOffsetDeg := 0.0;                        // 清偏置保持量（锁存量） / Clear offset
    IF _eState = E_DL_GpaState.eFault THEN
        _eState := E_DL_GpaState.eIdle;        // 故障相迁出：回未使能 / Fault exit to idle
    END_IF
END_IF
IF _bCfgBad THEN                               // 组态域闸 / Config gate
    _uFault := 16#0004_04A7;                   // 故障级：相位对齐故障总码 / Motion fault code
    _eCause := E_DL_GpaCause.eCfgIllegal;      // 归因：组态非法 / Cause: illegal config
    _bFault := TRUE;                           // 标志与码位配对（R45） / Flag paired with code
END_IF
IF (NOT _bFault) AND _bNonFin THEN             // 非有限锁存 / Non-finite latch
    _uFault := 16#0004_04A7;
    _eCause := E_DL_GpaCause.eNonFinite;       // 归因：非有限 / Cause: non-finite
    _bFault := TRUE;
END_IF

(* —— 段 3：偏置补偿（目标偏置 → 限幅 → 限速；仅无故障且未在窗时动作） —— *)
IF (NOT _bFault) AND (_eState = E_DL_GpaState.eAlign) AND (NOT _bInPhase) THEN
    _fCmdDeg := -_fErrDeg * fGainDegPerDeg;                    // 反向补偿目标 / Target compensation
    IF _fCmdDeg > fOffsetMaxDeg THEN                           // 偏置上限钳制 / Offset high clamp
        _fCmdDeg := fOffsetMaxDeg;
    ELSIF _fCmdDeg < -fOffsetMaxDeg THEN                       // 偏置下限钳制 / Offset low clamp
        _fCmdDeg := -fOffsetMaxDeg;
    END_IF
    IF (_fCmdDeg - _fOffsetDeg) > fOffsetStepDeg THEN          // 向上限速 / Upward rate limit
        _fOffsetDeg := _fOffsetDeg + fOffsetStepDeg;
    ELSIF (_fOffsetDeg - _fCmdDeg) > fOffsetStepDeg THEN       // 向下限速 / Downward rate limit
        _fOffsetDeg := _fOffsetDeg - fOffsetStepDeg;
    ELSE
        _fOffsetDeg := _fCmdDeg;                               // 直接跟随 / Follow target
    END_IF
    IF _fOffsetDeg > fOffsetMaxDeg THEN                        // 限速后二次复核上限 / Post-limit high
        _fOffsetDeg := fOffsetMaxDeg;
    ELSIF _fOffsetDeg < -fOffsetMaxDeg THEN                    // 限速后二次复核下限 / Post-limit low
        _fOffsetDeg := -fOffsetMaxDeg;
    END_IF
END_IF

(* —— 段 4：故障解除式（R240；全当拍量）：rtReset.Q / NOT _bCfgBad / NOT _bNonFin —— *)
IF rtReset.Q AND (NOT _bCfgBad) AND (NOT _bNonFin) THEN
    _bFault := FALSE;                          // 清故障锁存位（锁存量） / Clear fault latch
    _uFault := 16#0000_0000;                   // 清故障锁存码（锁存量） / Clear fault code
    _eCause := E_DL_GpaCause.eNone;            // 清成因（锁存量） / Clear cause
END_IF

(* —— 段 4A：故障锁存相位迁移闸（偏置冻结保持） —— *)
IF _bFault AND (_eState <> E_DL_GpaState.eFault) THEN
    _eState := E_DL_GpaState.eFault;           // 锁存即入故障相 / Latch enters fault phase
END_IF

(* —— 段 5：相位机（CASE 全覆盖 + ELSE 兜底） —— *)
CASE _eState OF

E_DL_GpaState.eIdle:
    IF bEnable AND (NOT _bFault) THEN          // 使能条件 / Enable gate
        _fOffsetDeg := 0.0;                    // 起始偏置清零（无扰） / Reset offset on start
        _eState := E_DL_GpaState.eAlign;       // 进对齐相 / Enter alignment
    END_IF

E_DL_GpaState.eAlign:
    IF _bInPhase THEN                          // 出口 1：相位在窗 / In phase
        _eState := E_DL_GpaState.eReady;       // 进可啮合相 / Enter ready
    ELSIF NOT bEnable THEN                     // 出口 2：撤使能（前置消失） / Disable
        _eState := E_DL_GpaState.eIdle;
    END_IF

E_DL_GpaState.eReady:
    IF NOT _bInPhase THEN                      // 相位漂出窗口：回对齐相 / Phase drifted out
        _eState := E_DL_GpaState.eAlign;
    ELSIF NOT bEnable THEN                     // 撤使能：回未使能 / Disable returns idle
        _eState := E_DL_GpaState.eIdle;
    END_IF

E_DL_GpaState.eFault:
    ;                                          // 故障相：偏置冻结，仅段 4 复位沿可迁出 / Frozen, reset only

ELSE
    _uFault := 16#0004_04A7;                   // 故障级：非法相位兜底（归并总码） / Illegal phase fallback
    _eCause := E_DL_GpaCause.eCfgIllegal;      // 归因：相位非法归并组态 / Cause: phase illegal
    _bFault := TRUE;
    _eState := E_DL_GpaState.eFault;           // 强制回故障相 / Force fault phase

END_CASE

(* —— 段 6：出口单点映射（名实同源；故障相偏置冻结、许可撤销） —— *)
IF _bFault THEN
    nErrId := _uFault;                         // 故障锁存码回放 / Replay latched code
    fPhaseErrDeg := 0.0;                       // 故障相相位差出口强制 0 / Error forced zero
    bInPhase := FALSE;                         // 故障相啮合许可强制撤销（安全侧） / Permit forced off
    fOffsetDeg := _fOffsetDeg;                 // 故障相偏置冻结保持 / Offset frozen
ELSE
    nErrId := 16#0000_0000;                    // 无故障：本件无信息码 / No fault, no info code
    fPhaseErrDeg := _fErrDeg;                  // 相位差出口 / Error outlet
    bInPhase := _bInPhase;                     // 啮合许可出口 / Permit outlet
    fOffsetDeg := _fOffsetDeg;                 // 偏置出口 / Offset outlet
END_IF
bError := _bFault;                             // 故障标志同源 / Flag from latch
eState := _eState;                             // 状态出口 / State outlet
eCause := _eCause;                             // 成因出口 / Cause outlet

END_FUNCTION_BLOCK

(* ---- FB_DL_HoneHeadExpansionSeq.st ---- *)
//==============================================================================
// 功能块：FB_DL_HoneHeadExpansionSeq ｜ 中文名称：珩磨头涨缩与往复联动序（复杂度 C4）
// 所属子库：DL_Motion ｜ 版本 VERSION: v1.0.0 ｜ 兼容：CODESYS V3.5+ / TwinCAT 3 / 汇川 InoProShop
// 功能描述：珩磨头按压力曲线涨开油石——接近 → 压力爬坡涨开 → 保压珩磨 → 缩回退刀
//           → 完成。涨开量 = 基准涨开量 + 油石磨损补偿（按件数线性累加）；压力闭环
//           用纯比例 + 死区（无积分器，杜绝饱和），指令按爬坡速率限幅；中止立即泄压、
//           压力降到安全值以下才允许退刀（禁止带压退刀）。
// 开源溯源 (Origin)：道莅原创实现（参考 ISO 12180 珩磨工艺与油石磨损补偿工程惯例
//           分类与参数域，许可证=MIT，借鉴点=「按件数线性补偿涨开量 + 定压保压」工艺序）
// 单位表：压力[bar] / 涨开量[μm] / 时间[ms] / 计数[件]
// 错误码表（Motion 段 0008，故障窗口 0B01~0B08，信息窗口 0B11）：
//   16#0008_0B01 故障级：组态非法（目标压/爬坡率/上限/时间量 <= 0，或磨损系数 < 0）
//   16#0008_0B02 故障级：压力反馈入口非有限（NaN / Inf）或幅值超合法上限，拒算
//   16#0008_0B03 故障级：涨开量 > fMaxExpandUm，拒动并置 xOverExpand
//   16#0008_0B04 故障级：涨开爬坡超时（压力未进入目标带宽）
//   16#0008_0B05 故障级：保压期压力跌出带宽（掉压）
//   16#0008_0B06 故障级：泄压超时（压力未降到安全值，禁止带压退刀）
//   16#0008_0B07 故障级：缩回超时（tRetractTime 满时压力仍高于安全值，退刀未完成）
//   16#0008_0B08 故障级兜底：状态机落 ELSE 非法态，全输出断
//   16#0008_0B11 信息级：涨缩循环完成（完成拍，不置 bError）
//           故障级码全部锁存回放（R187），唯一清除路径 = bReset 上升沿。
// 状态机：E_DL_HoneExpState（七态：eIdle=0 / eApproach=10 / eExpand=20 / eDwell=30 /
//           eRetract=40 / eDone=50 / eFault=99）。中止两段化不占相位，由内部段号
//           _uAbortStage 驱动（0 无 / 1 泄压中 / 2 退刀中）。
// 边界行为：① eApproach 为固定接近延时相，不设超时（无故障码，仅作换向让位）；② 涨开
//           与缩回两命令在段 10 互斥，任何相不得同时置位；③ 带压退刀被物理禁止：中止段
//           A 只泄压不退刀，压力降到 DL_HNE_SAFE_BAR 以下才进段 B；④ 保压期压力跌出带宽
//           持续 DL_HNE_DROP_T 即锁存 0B05，不用单拍瞬时值；⑤ 七态 CASE 每态显式 +
//           ELSE 兜底 → 0B08 全断。
// 语义假设：① 压力指令为 bar 量纲的比例阀指令，0 bar = 泄压；② 涨开量与压力非线性对
//           应，故涨开量只作磨损补偿核算（fExpandUm 供上层显示与上限校验），不参与压力
//           闭环；③ 闭环执行周期按 DL_HNE_DT_S 假定 10 ms，本件无任务周期引脚，故以常量
//           声明该假定，换平台须同步。
// 依赖纪律：仅 Standard.library（TON / R_TRIG）；零 GVL、零 VAR_EXTERNAL、零物理地址。
// 修订历史：v1.0.0 2026-11-25 R88 首版（无人值守批次 · 复杂件 C4 · 序号 2）
//==============================================================================

(*------------------------------------------------------------------------------
 * 枚举: E_DL_HoneExpState（归属本功能块，同文件发布，全库唯一定义）
 * 含义: 珩磨头涨缩相位，与段 9 状态机、段 10 输出置位一一对应。
 *-----------------------------------------------------------------------------*)
TYPE E_DL_HoneExpState :
(
    eIdle     := 0,  // 空闲：等启动沿 / Idle, awaiting the start edge
    eApproach := 10, // 接近：固定延时让位，为涨开做准备 / Approach, fixed delay before expansion
    eExpand   := 20, // 涨开：压力按爬坡率升到目标带宽 / Expand, pressure ramps into the target band
    eDwell    := 30, // 保压：定压珩磨计时，监视掉压 / Dwell, timed honing with drop monitoring
    eRetract  := 40, // 缩回：压力归零并缩回退刀 / Retract, pressure zeroed before withdrawal
    eDone     := 50, // 完成：本件循环结束 / Done, the cycle finished
    eFault    := 99  // 故障：组态/掉压/超时/非法态 / Fault, configuration, pressure drop, timeout or illegal state
);
END_TYPE

FUNCTION_BLOCK FB_DL_HoneHeadExpansionSeq
VAR_INPUT
    xEnable          : BOOL;   // 使能，FALSE 期间按中止处理 [—] / Enable, a drop is treated as an abort
    xStart           : BOOL;   // 启动请求，上升沿生效 [—] / Start request, rising edge effective
    xAbort           : BOOL;   // 中止请求，任意拍生效（立即泄压） [—] / Abort request, effective on any scan
    xReset           : BOOL;   // 故障复位，上升沿清全部锁存 [—] / Fault reset, rising edge clears all latches
    fTargetPressBar  : LREAL;  // 目标珩磨压力 [bar]，须 > 0 / Target honing pressure [bar], must be > 0
    fPressFbBar      : LREAL;  // 压力实际反馈 [bar] / Actual pressure feedback [bar]
    fRampRateBarPerS : LREAL;  // 压力指令爬坡速率 [bar/s]，须 > 0 / Command ramp rate [bar/s], must be > 0
    tDwellTime       : TIME;   // 保压珩磨时长 [ms] / Dwell honing time [ms]
    tRetractTime     : TIME;   // 缩回退刀时长 [ms] / Retract time [ms]
    fStoneWearUmPerPc: LREAL;  // 油石每件磨损量 [μm/件] / Stone wear per piece [um/pc]
    nPieceCount      : UDINT;  // 累计加工件数 [件]，用于磨损补偿 / Accumulated piece count for wear compensation
    fMaxExpandUm     : LREAL;  // 涨开量上限 [μm]，须 > 0 / Expansion ceiling [um], must be > 0
    tPressTimeout    : TIME;   // 涨开爬坡与泄压超时 [ms] / Ramp and vent timeout [ms]
END_VAR
VAR_OUTPUT
    fPressCmdBar     : LREAL;  // 压力指令出口 [bar]，0 = 泄压 / Pressure command outlet [bar], 0 = vented
    xExpandCmd       : BOOL;   // 涨开命令（油石外张） [—] / Expansion command
    xRetractCmd      : BOOL;   // 缩回命令（油石内收退刀） [—] / Retract command
    bRunning         : BOOL;   // 循环运行中（非空闲非完成非故障非中止） [—] / Cycle active
    bDone            : BOOL;   // 单件循环完成相电平 [—] / Cycle done, level in the done phase
    bError           : BOOL;   // 故障级标志，仅故障级码置位 [—] / Fault-class flag, fault-level codes only
    nErrCode         : UDINT;  // 错误码，0 = 无错 [—] / Error code, 0 = none
    fExpandUm        : LREAL;  // 涨开量出口 [μm] = 基准 + 磨损补偿 / Expansion outlet [um] = base plus wear
    fWearCompUm      : LREAL;  // 磨损补偿量出口 [μm] = 每件磨损 × 件数 / Wear compensation outlet [um]
    xOverExpand      : BOOL;   // 涨开量超上限（拒动锁存） [—] / Expansion beyond the ceiling, latched
END_VAR
VAR
    _eState          : E_DL_HoneExpState := E_DL_HoneExpState.eIdle; // 当前相位 [—] / Current phase
    _bInit           : BOOL := FALSE;   // 首扫标志，取非判定 [—] / First-scan flag, tested negated
    _fPressCmd       : LREAL;           // 压力指令保持量（速率限幅后） [bar] / Held command after rate limiting [bar]
    _fWearCompUm     : LREAL;           // 内部磨损补偿量 [μm] / Internal wear compensation [um]
    _fExpandUm       : LREAL;           // 内部涨开量 [μm] / Internal expansion [um]
    _bCfgBad         : BOOL;            // 组态非法锁存 / Illegal configuration latch
    _bCfgOk          : BOOL;            // 本拍组态合法（派生量不锁存） [—] / Configuration legal this scan, derived
    _bSigBad         : BOOL;            // 压力反馈非有限锁存 / Non-finite pressure feedback latch
    _bOverExpand     : BOOL;            // 涨开量超上限锁存 / Over-expansion latch
    _bRampTmo        : BOOL;            // 涨开爬坡超时锁存 / Ramp timeout latch
    _bDropErr        : BOOL;            // 保压掉压锁存 / Pressure drop latch
    _bVentTmo        : BOOL;            // 泄压超时锁存 / Vent timeout latch
    _bRetractTmo     : BOOL;            // 缩回超时锁存 / Retract timeout latch
    _bIllegal        : BOOL;            // 非法状态标志 / Illegal state flag
    _bInfoDone       : BOOL;            // 循环完成信息当拍标志 / Cycle-done info flag of this scan
    _bAbortReq       : BOOL;            // 中止请求合成（xAbort 或失能） [—] / Combined abort request
    _bBandOk         : BOOL;            // 压力在目标带宽内（派生量） [—] / Pressure inside the target band, derived
    _bSafePressure   : BOOL;            // 压力已降到安全值以下（派生量） [—] / Pressure below the safe value, derived
    _uAbortStage     : UINT;            // 中止段号 0=无 1=泄压中 2=退刀中 / Abort stage 0 none 1 venting 2 retracting
    rtStart          : R_TRIG;          // 启动沿，段 7 无条件刷新 [—] / Start edge, refreshed in segment 7
    rtReset          : R_TRIG;          // 复位沿，段 7 无条件刷新 [—] / Reset edge, refreshed in segment 7
    tonApproach      : TON;             // 接近让位延时 [ms] / Approach delay [ms]
    tonRamp          : TON;             // 涨开爬坡超时 [ms] / Ramp timeout [ms]
    tonDwell         : TON;             // 保压珩磨计时 [ms] / Dwell honing timer [ms]
    tonPressDrop     : TON;             // 保压掉压持续窗 [ms] / Pressure-drop persistence window [ms]
    tonRetract       : TON;             // 缩回退刀计时 [ms] / Retract timer [ms]
    tonVent          : TON;             // 中止泄压超时 [ms] / Abort venting timeout [ms]
    tonAbortRetract  : TON;             // 中止退刀计时 [ms] / Abort retract timer [ms]
END_VAR
VAR_TEMP
    fErr             : LREAL;           // 本拍压力偏差暂存 [bar] / Pressure error scratch of this scan [bar]
    fDes             : LREAL;           // 本拍期望指令暂存 [bar] / Desired command scratch of this scan [bar]
    fRampStep        : LREAL;           // 本拍允许变化量暂存 [bar] / Allowed change per scan [bar]
END_VAR
VAR CONSTANT
    DL_EPS            : LREAL := 1.0E-9;     // 浮点容差零点，兼作除法分母下限 / Float epsilon, also the divisor floor
    DL_HNE_DT_S       : LREAL := 0.01;       // 闭环假定执行周期 [s]（10 ms 任务） / Assumed control period [s]
    DL_HNE_KP         : LREAL := 2.0;        // 压力闭环比例增益 [bar/bar] / Proportional gain [bar/bar]
    DL_HNE_DEAD_BAR   : LREAL := 0.05;       // 比例控制死区 [bar]，死区内保持指令 / Proportional dead band [bar]
    DL_HNE_BAND_RATIO : LREAL := 0.10;       // 目标带宽比例项 [倍] / Target band ratio term
    DL_HNE_BAND_MIN   : LREAL := 0.50;       // 目标带宽最小绝对值 [bar] / Minimum absolute band [bar]
    DL_HNE_BASE_UM    : LREAL := 25.0;       // 油石基准涨开量 [μm] / Base stone expansion [um]
    DL_HNE_CMD_MAX    : LREAL := 60.0;       // 压力指令幅值上限 [bar] / Command magnitude ceiling [bar]
    DL_HNE_SAFE_BAR   : LREAL := 0.50;       // 退刀前压力安全值 [bar] / Safe pressure before retraction [bar]
    DL_HNE_PRESS_MAX  : LREAL := 400.0;      // 压力反馈合法幅值上限 [bar] / Legal feedback ceiling [bar]
    DL_HNE_APPROACH_T : TIME  := T#800MS;    // 接近让位固定延时 [ms] / Fixed approach delay [ms]
    DL_HNE_DROP_T     : TIME  := T#300MS;    // 掉压持续判定窗 [ms] / Drop persistence window [ms]
END_VAR

(*------------------------------------------------------------------------------
 * 段 1｜每拍预置：全部输出先落安全侧，单拍标志预清零
 *      All outputs preset to the safe side, one-shot flags pre-cleared
 *-----------------------------------------------------------------------------*)
fPressCmdBar := 0.0;                        // 压力指令先归零（泄压安全侧） / Command zeroed, vented side
xExpandCmd := FALSE; xRetractCmd := FALSE;  // 涨开/缩回命令先断 / Expansion and retract commands cleared
bRunning := FALSE;  bDone := FALSE;         // 运行与完成标志每拍重算 / Running and done flags recomputed
bError := FALSE;    nErrCode := 16#0000_0000; // 故障标志与错误码每拍重算 / Fault flag and code recomputed
xOverExpand := FALSE;                       // 超涨开标志每拍重算 / Over-expansion flag recomputed
_bIllegal := FALSE; _bInfoDone := FALSE;    // 非法态与完成信息预清零 / Illegal and done-info flags pre-cleared

(*------------------------------------------------------------------------------
 * 段 2｜首扫初始化：相位、指令保持量与中止段号复位
 *      First-scan initialisation of phase, held command and abort stage
 *-----------------------------------------------------------------------------*)
IF NOT _bInit THEN
    _eState      := E_DL_HoneExpState.eIdle; // 相位从空闲起步 / Phase starts idle
    _fPressCmd := 0.0;  _fWearCompUm := 0.0; _fExpandUm := 0.0; // 指令/磨损/涨开量从零起步 / Command, wear and expansion at zero
    _uAbortStage := 0;                       // 中止段号从零起步 / Abort stage starts at zero
    _bInit       := TRUE;                    // 首扫只做一次 / The first scan runs once
END_IF

(*------------------------------------------------------------------------------
 * 段 3｜入口非有限闸 + 组态闸（浮点量逐只双侧幅值判，时间量下限判）
 *      Non-finite inlet gate and configuration gates
 *-----------------------------------------------------------------------------*)
IF NOT (fPressFbBar > -1.0E30 AND fPressFbBar < 1.0E30) THEN _bSigBad := TRUE; END_IF    // 压力反馈非有限 → 0B02 / Non-finite feedback, 0B02
IF ABS(fPressFbBar) > DL_HNE_PRESS_MAX THEN _bSigBad := TRUE; END_IF                   // 反馈幅值超上限 → 0B02 / Beyond the ceiling, 0B02
IF NOT (fTargetPressBar > -1.0E30 AND fTargetPressBar < 1.0E30) THEN _bCfgBad := TRUE; END_IF // 目标压非有限 → 0B01 / Non-finite target, 0B01
IF NOT (fRampRateBarPerS > -1.0E30 AND fRampRateBarPerS < 1.0E30) THEN _bCfgBad := TRUE; END_IF // 爬坡率非有限 → 0B01 / Non-finite ramp, 0B01
IF NOT (fMaxExpandUm > -1.0E30 AND fMaxExpandUm < 1.0E30) THEN _bCfgBad := TRUE; END_IF  // 涨开上限非有限 → 0B01 / Non-finite ceiling, 0B01
IF NOT (fStoneWearUmPerPc > -1.0E30 AND fStoneWearUmPerPc < 1.0E30) THEN _bCfgBad := TRUE; END_IF // 磨损系数非有限 → 0B01 / Non-finite wear, 0B01
IF (fTargetPressBar <= DL_EPS) OR (fRampRateBarPerS <= DL_EPS) OR (fMaxExpandUm <= DL_EPS)
   OR (fStoneWearUmPerPc < 0.0) THEN _bCfgBad := TRUE; END_IF // 三者须为正且磨损非负 → 0B01 / Positive values required, 0B01
IF (tDwellTime <= T#0MS) OR (tRetractTime <= T#0MS) OR (tPressTimeout <= T#0MS) THEN _bCfgBad := TRUE; END_IF // 时间量须为正 → 0B01 / Time values must be positive
_bCfgOk := NOT _bCfgBad;                    // 本拍组态合法派生量 / Configuration-legal derived flag of this scan

(*------------------------------------------------------------------------------
 * 段 4｜磨损补偿与涨开量核算 + 超涨开拒动判定
 *      Wear compensation, expansion accounting and the over-expansion check
 *-----------------------------------------------------------------------------*)
_fWearCompUm := fStoneWearUmPerPc * UDINT_TO_LREAL(nPieceCount); // 磨损补偿 [μm] = 每件磨损 × 件数 / Wear = per-piece wear times pieces
_fExpandUm   := DL_HNE_BASE_UM + _fWearCompUm;                   // 涨开量 [μm] = 基准 + 磨损补偿 / Expansion = base plus wear
IF (_bCfgOk) AND (_fExpandUm > fMaxExpandUm) THEN
    _bOverExpand := TRUE;                   // 涨开量超上限，拒动锁存 → 0B03 / Beyond the ceiling, code 0B03
END_IF
fWearCompUm := _fWearCompUm; fExpandUm := _fExpandUm; // 磨损补偿与涨开量出口 [μm] / Wear and expansion outlets [um]
xOverExpand := _bOverExpand;                // 超涨开出口 [—] / Over-expansion outlet

(*------------------------------------------------------------------------------
 * 段 5｜压力闭环（纯比例 + 死区，无积分器）+ 爬坡速率限幅
 *      Pressure loop, proportional only with a dead band, plus ramp rate limiting
 *-----------------------------------------------------------------------------*)
IF ((_eState = E_DL_HoneExpState.eExpand) OR (_eState = E_DL_HoneExpState.eDwell))
   AND (_uAbortStage = 0) AND (NOT _bCfgBad) AND (NOT _bSigBad) THEN
    fErr := fTargetPressBar - fPressFbBar;  // 压力偏差 [bar] / Pressure error [bar]
    IF ABS(fErr) > DL_HNE_DEAD_BAR THEN
        fDes := _fPressCmd + DL_HNE_KP * fErr; // 比例增量，死区外才动 / Proportional increment outside the dead band
    ELSE
        fDes := _fPressCmd;                 // 死区内保持（无积分器，杜绝饱和） / Held inside the dead band, no integrator
    END_IF
    IF fDes < 0.0 THEN fDes := 0.0; END_IF  // 指令下钳 0（不吸真空） / Lower clamp at zero
    IF fDes > DL_HNE_CMD_MAX THEN fDes := DL_HNE_CMD_MAX; END_IF // 指令上钳幅值上限 / Upper clamp at the ceiling
    fRampStep := fRampRateBarPerS * DL_HNE_DT_S; // 本拍允许变化量 [bar] / Allowed change per scan [bar]
    IF (fDes - _fPressCmd) > fRampStep THEN fDes := _fPressCmd + fRampStep;      // 正向限幅 / Positive ramp limit
    ELSIF (fDes - _fPressCmd) < (0.0 - fRampStep) THEN fDes := _fPressCmd - fRampStep; // 反向限幅 / Negative ramp limit
    END_IF
    _fPressCmd := fDes;                     // 指令保持量推进 / Held command advanced
ELSE
    _fPressCmd := 0.0;                      // 非涨开相一律归零（泄压） / Zeroed outside the expansion phases
END_IF
fPressCmdBar := _fPressCmd;                 // 压力指令出口 [bar] / Pressure command outlet [bar]
_bBandOk := ABS(fPressFbBar - fTargetPressBar) <= (fTargetPressBar * DL_HNE_BAND_RATIO + DL_HNE_BAND_MIN); // 带宽判据 / Band criterion
_bSafePressure := fPressFbBar <= DL_HNE_SAFE_BAR;  // 安全压判据（退刀许可） / Safe-pressure criterion for retraction

(*------------------------------------------------------------------------------
 * 段 6｜中止入口（段 0→1，立即泄压）与复位
 *      Abort entry, immediate venting, and the reset edge
 *-----------------------------------------------------------------------------*)
_bAbortReq := xAbort OR (NOT xEnable);      // 中止请求合成：显式中止或失能 / Combined abort: explicit abort or enable loss
IF _bAbortReq AND (_uAbortStage = 0) AND (_eState <> E_DL_HoneExpState.eIdle)
   AND (_eState <> E_DL_HoneExpState.eDone) AND (_eState <> E_DL_HoneExpState.eFault) THEN
    _uAbortStage := 1;                      // 进中止段 A：立即泄压，禁带压退刀 / Enter abort stage A, vent first
END_IF
IF rtReset.Q THEN
    _bCfgBad := FALSE;  _bSigBad := FALSE;  _bOverExpand := FALSE; // 复位清组态/反馈/超涨开锁存 / Clears configuration, feedback, expansion
    _bRampTmo := FALSE; _bDropErr := FALSE; _bVentTmo := FALSE; _bRetractTmo := FALSE; // 复位清爬坡/掉压/泄压/缩回锁存 / Clears ramp, drop, vent, retract
END_IF

(*------------------------------------------------------------------------------
 * 段 7｜定时器与边沿无条件周期刷新（R7：CASE 之外每拍必调，各司其职不复用）
 *      Timers and edges refreshed unconditionally every scan, outside the CASE
 *-----------------------------------------------------------------------------*)
rtStart(CLK := xStart); rtReset(CLK := xReset); // 启动沿与复位沿无条件刷新 / Start and reset edges refreshed
tonApproach(IN := (_eState = E_DL_HoneExpState.eApproach) AND (_uAbortStage = 0), PT := DL_HNE_APPROACH_T); // 接近让位延时 / Approach delay
tonRamp(IN := (_eState = E_DL_HoneExpState.eExpand) AND (_uAbortStage = 0), PT := tPressTimeout);            // 涨开爬坡超时 / Ramp timeout
tonDwell(IN := (_eState = E_DL_HoneExpState.eDwell) AND (_uAbortStage = 0), PT := tDwellTime);               // 保压计时 / Dwell timer
tonPressDrop(IN := (_eState = E_DL_HoneExpState.eDwell) AND (NOT _bBandOk), PT := DL_HNE_DROP_T);            // 掉压持续窗 / Drop window
tonRetract(IN := (_eState = E_DL_HoneExpState.eRetract) AND (_uAbortStage = 0), PT := tRetractTime);         // 缩回计时 / Retract timer
tonVent(IN := (_uAbortStage = 1), PT := tPressTimeout);                                                      // 中止泄压超时 / Abort vent timeout
tonAbortRetract(IN := (_uAbortStage = 2), PT := tRetractTime);                                               // 中止退刀计时 / Abort retract timer

(*------------------------------------------------------------------------------
 * 段 8｜中止段推进（1 泄压 → 压力安全值以下才进 2 退刀 → 收口）
 *      Abort progression, retraction only after the pressure is below the safe value
 *-----------------------------------------------------------------------------*)
IF (_uAbortStage = 1) AND _bSafePressure THEN
    _uAbortStage := 2;                      // 压力已泄到安全值，进退刀段 / Pressure safe, enter retraction
ELSIF (_uAbortStage = 1) AND tonVent.Q THEN
    _bVentTmo := TRUE; _uAbortStage := 0;   // 泄压超时，禁止带压退刀 → 0B06 / Vent timeout, 0B06
    _eState   := E_DL_HoneExpState.eFault;  // 落故障 / Fall to fault
END_IF
IF (_uAbortStage = 2) AND tonAbortRetract.Q THEN
    _uAbortStage := 0;                      // 退刀完成，中止收口 / Retraction done, abort closed
    _eState      := E_DL_HoneExpState.eIdle; // 回空闲 / Back to idle
END_IF
(*------------------------------------------------------------------------------
 * 段 9｜状态机（中止期间迁移冻结；本段只做迁移，输出在段 10）
 *      Phase machine, transitions frozen while aborting, outputs in segment 10
 *-----------------------------------------------------------------------------*)
IF _uAbortStage = 0 THEN
    CASE _eState OF
        E_DL_HoneExpState.eIdle:            // 空闲：启动沿 + 组态合法 + 未超涨开才进接近 / Idle, legal start edge only
            IF rtStart.Q AND _bCfgOk AND (NOT _bSigBad) AND (NOT _bOverExpand) AND (NOT _bAbortReq) THEN
                _fPressCmd := 0.0;          // 新循环指令复位 / Command reset for the new cycle
                _eState    := E_DL_HoneExpState.eApproach; // 进接近相 / To the approach phase
            END_IF
        E_DL_HoneExpState.eApproach:        // 接近：固定让位延时满即涨开 / Approach, expansion after the fixed delay
            IF tonApproach.Q THEN _eState := E_DL_HoneExpState.eExpand; END_IF // 延时满，进涨开相 / Delay elapsed, expand
        E_DL_HoneExpState.eExpand:          // 涨开：压力进入带宽即进保压，超时落故障 / Expand into the band or time out
            IF _bBandOk THEN _eState := E_DL_HoneExpState.eDwell; // 压力进带宽，进保压相 / In band, to dwell
            ELSIF tonRamp.Q THEN _bRampTmo := TRUE; _eState := E_DL_HoneExpState.eFault; // 爬坡超时 → 0B04 / Ramp timeout, 0B04
            END_IF
        E_DL_HoneExpState.eDwell:           // 保压：掉压超窗落故障，计时满进缩回 / Dwell, drop faults, timer to retract
            IF tonPressDrop.Q THEN _bDropErr := TRUE; _eState := E_DL_HoneExpState.eFault; // 掉压持续 → 0B05 / Pressure drop, 0B05
            ELSIF tonDwell.Q THEN _eState := E_DL_HoneExpState.eRetract; // 保压满，进缩回相 / Dwell elapsed, retract
            END_IF
        E_DL_HoneExpState.eRetract:         // 缩回：退刀计时满且压力已安全才完成 / Retract done once timed and safe
            IF tonRetract.Q AND (NOT _bSafePressure) THEN
                _bRetractTmo := TRUE; _eState := E_DL_HoneExpState.eFault; // 计时满仍带压 → 0B07 / Still pressurized, 0B07
            ELSIF tonRetract.Q THEN
                _bInfoDone := TRUE;         // 置循环完成信息 / Raise the cycle-done info
                _eState    := E_DL_HoneExpState.eDone; // 进完成相 / To the done phase
            END_IF
        E_DL_HoneExpState.eDone:            // 完成：启动撤销且无中止请求才回空闲 / Done, back to idle once start drops
            IF (NOT xStart) AND (NOT _bAbortReq) THEN _eState := E_DL_HoneExpState.eIdle; END_IF
        E_DL_HoneExpState.eFault:           // 故障：复位沿且组态合法且未超涨开才回空闲 / Fault, reset edge only
            IF rtReset.Q AND _bCfgOk AND (NOT _bSigBad) AND (NOT _bOverExpand) THEN _eState := E_DL_HoneExpState.eIdle; END_IF
        ELSE                                // 非法状态兜底（R6：CASE 必带 ELSE）/ Illegal-state fallback
            _bIllegal := TRUE; _eState := E_DL_HoneExpState.eFault; // 非法态 → 0B08，落故障 / Illegal state, 0B08
    END_CASE
END_IF
(*------------------------------------------------------------------------------
 * 段 10｜输出置位（涨开与缩回互斥；中止段 A 只泄压不退刀）
 *      Output assignment, expand and retract exclusive, abort stage A vents only
 *-----------------------------------------------------------------------------*)
xExpandCmd := FALSE;                        // 默认两命令先断，再由状态判定置位（R88 修复：原 CASE ELSE 覆盖涨开命令） / default both off (R88 fix)
xRetractCmd := FALSE;                       // 缩回命令默认断 / retract default off
IF (_eState = E_DL_HoneExpState.eExpand) OR (_eState = E_DL_HoneExpState.eDwell) THEN
    xExpandCmd := TRUE;                     // 涨开相与保压相：油石外张 / Expand and dwell, stone outwards
END_IF
CASE _eState OF
    E_DL_HoneExpState.eRetract:             // 缩回相：油石内收退刀 / Retract phase, stone inwards
        xRetractCmd := TRUE;                // 缩回命令 / Retract command
    E_DL_HoneExpState.eDone:                // 完成相：完成电平 / Done phase, done level
        bDone := TRUE;                      // 循环完成 / Cycle done
    ELSE
        xRetractCmd := FALSE;               // 兜底：仅保持缩回断，涨开指令由上方状态判定决定，不得覆盖 / fallback keeps retract off only
END_CASE
IF _uAbortStage >= 1 THEN
    xExpandCmd := FALSE;                    // 中止段 A：涨开命令立即断 / Abort A, expansion cut immediately
    fPressCmdBar := 0.0;                    // 立即泄压（泄压优先于一切） / Vent immediately, before anything else
    xRetractCmd := (_uAbortStage = 2);      // 压力已安全才退刀，禁带压退刀 / Retract only once the pressure is safe
END_IF
bRunning := (_eState <> E_DL_HoneExpState.eIdle) AND (_eState <> E_DL_HoneExpState.eDone)
            AND (_eState <> E_DL_HoneExpState.eFault) AND (_uAbortStage = 0); // 运行标志 / Running flag

(*------------------------------------------------------------------------------
 * 段 11｜错误码映射（锁存回放，R187：故障相不按当下输入重推断）
 *      Error-code map, latched replay
 *-----------------------------------------------------------------------------*)
IF _bIllegal THEN nErrCode := 16#0008_0B08; bError := TRUE;        // 故障级兜底：非法态 / Fault, illegal state fallback
ELSIF _bCfgBad THEN nErrCode := 16#0008_0B01; bError := TRUE;      // 故障级：组态非法 / Fault, illegal configuration
ELSIF _bSigBad THEN nErrCode := 16#0008_0B02; bError := TRUE;      // 故障级：压力反馈非有限 / Fault, non-finite feedback
ELSIF _bOverExpand THEN nErrCode := 16#0008_0B03; bError := TRUE;  // 故障级：涨开量超上限 / Fault, over expansion
ELSIF _bRampTmo THEN nErrCode := 16#0008_0B04; bError := TRUE;     // 故障级：涨开爬坡超时 / Fault, ramp timeout
ELSIF _bDropErr THEN nErrCode := 16#0008_0B05; bError := TRUE;     // 故障级：保压掉压 / Fault, pressure drop
ELSIF _bVentTmo THEN nErrCode := 16#0008_0B06; bError := TRUE;     // 故障级：泄压超时/带压退刀 / Fault, vent timeout
ELSIF _bRetractTmo THEN nErrCode := 16#0008_0B07; bError := TRUE;  // 故障级：缩回超时 / Fault, retract timeout
ELSIF _bInfoDone THEN nErrCode := 16#0008_0B11;                    // 信息级：循环完成，不置 bError / Info, cycle done
END_IF
END_FUNCTION_BLOCK

(* ---- FB_DL_LabelApplySync.st ---- *)
//==============================================================================
// 功能块：FB_DL_LabelApplySync ｜ 中文名称：贴标同步出标控制
// 所属子库：DL_Motion ｜ 版本：v1.0.0 ｜ 兼容：CODESYS V3.5+ / TwinCAT 3 / 汇川 InoProShop
// 功能描述：卷料贴标机的出标同步件。编码器累计脉冲差分求卷材位移（差分按带符号减法，
//           32 位回绕时符号自然正确，禁止按绝对值比较），按标签节距分频出标扳机，扣
//           除出标提前量，并给出相位误差、线速度与低速禁止出标判据。低速时相位估算不
//           可靠，硬出标会贴歪，故低速一律抑制出标并提示。本件只输出出标扳机与诊断
//           量，不改轴状态、不发运动指令（轴状态唯一属主是运动层，T1-6 纪律），也不
//           驱动贴标头气缸与真空（执行器归设备层）。
// 开源溯源 (Origin)：道莅原创实现（参考 公开工程惯例 分类与参数域）
// 单位表：累计脉冲[脉冲] / 脉冲当量[脉冲每毫米] / 节距与提前量[mm] / 线速度[米每分] /
//         相位误差[mm] / 触发脉宽[ms] / 扫描间隔[ms] / 出标计数[张]
// 错误码表：16#0004_01ED 信息级（提前量超一个节距被饱和钳位，钳到节距，不置 bError）/
//           16#0004_01EE 信息级（编码器低速，相位估算不可靠，暂停出标，不置 bError）/
//           16#0004_030F 故障级（脉冲当量或标签节距组态非法，置 bError，先判后除）/
//           16#0004_0310 故障级（输入非有限，置 bError）/ 16#0004_0311 故障级兜底
//           （状态机落 ELSE 非法状态，置 bError）。码位 16#0004 段，不越段不挪预留槽。
// 状态机：E_DL_LabelSyncState（eIdle=0 失能/待机 / eSync=10 同步出标 / eLowSpeed=20
//           低速抑制出标 / eFault=99 故障兜底），CASE 含 ELSE 兜底，ELSE 置 0311 并撤
//           出标扳机与许可。
// 边界行为：① 脉冲差分 nDelta := nNow − nPrev（DINT 回绕安全；上电首拍以当前脉冲为
//           基准，避免首拍巨量假位移）；② fPulsePerMm <= 0 或 fLabelPitchMm <= 0 → 故障
//           030F，全部除法位于该闸之后（先判后除）；③ 线速度低于 fSpeedMinMpm → 不出
//           标 + 信息 01EE + bLowSpeed，相位继续累计（回速后按相位补出，不丢位置）；
//           ④ 提前量超一个节距 → 钳到节距 + 信息 01ED；⑤ bLabelPresent := FALSE → 不出
//           标且 bMissedLabel 锁存（漏标次数由上层按本标志上升沿自行计数，本件不设死
//           计数器）；⑥ 失能 → bFireTrigger := FALSE + bValid := FALSE（R72）；⑦ 非有限
//           或解算溢出（NaN 自反判 + Inf 幅值上限判）→ 故障 0310，扳机撤。
// 修订历史：v1.0.0 2026-11-17 首版（R25 派单 · §4.13）
//==============================================================================
(*------------------------------------------------------------------------------
 * 枚举: E_DL_LabelSyncState（归属 DL_Motion，与 FB_DL_LabelApplySync 同文件）
 *----------------------------------------------------------------------------*)
TYPE E_DL_LabelSyncState :
(
    eIdle     := 0,   // 失能/待机：扳机撤，相位基准重新对齐 / Disabled, trigger dropped, phase re-based
    eSync     := 10,  // 同步出标：线速度达标，按节距分频出标 / Synchronised firing at the label pitch
    eLowSpeed := 20,  // 低速抑制：速度低于下限，不出标只累计相位 / Low speed, firing suppressed, phase still accumulated
    eFault    := 99   // 故障兜底：组态非法/非有限/非法状态 / Fault fallback
);
END_TYPE

(*==============================================================================
 * 功能块: FB_DL_LabelApplySync
 * 调用约定: 每个扫描周期无条件调用一次；nEncoderPulse 由高速计数或编码器模块刷新，
 *           uDeltaTimeMs 必须注入真实任务间隔。
 *============================================================================*)
FUNCTION_BLOCK FB_DL_LabelApplySync
VAR_INPUT
    nEncoderPulse  : DINT;                        // 编码器累计脉冲 [脉冲]，允许 32 位回绕 / Encoder accumulated pulses [pulse], 32-bit wrap allowed
    fPulsePerMm    : LREAL := 100.0;              // 脉冲当量 [脉冲每毫米]，须 > 0 / Pulse equivalent [pulse per mm], must be > 0
    fLabelPitchMm  : LREAL := 50.0;               // 标签节距 [mm]，须 > 0 / Label pitch [mm], must be > 0
    fLeadMm        : LREAL := 2.0;                // 出标提前量 [mm]，超一个节距被钳位 / Label lead [mm], clamped to one pitch
    fSpeedMinMpm   : LREAL := 5.0;                // 最低同步线速度 [米每分] / Minimum synchronised web speed [m per min]
    bLabelPresent  : BOOL;                        // 标签在位（缺标检测）/ Label present, missing-label detection
    tTriggerHold   : TIME := T#20MS;              // 出标触发脉宽 [ms] / Trigger pulse width [ms]
    uDeltaTimeMs   : UDINT;                       // 扫描间隔 [ms]，调用方注入，禁系统时间函数 / Scan interval [ms], caller-injected
    bEnable        : BOOL;                        // 总使能 / Master enable
    bReset         : BOOL;                        // 复位，上升沿清漏标/饱和提示/故障与计数 / Reset, rising edge clears the missed-label latch, hints, fault and counter
END_VAR
VAR_OUTPUT
    bFireTrigger   : BOOL;                        // 出标触发（脉宽 tTriggerHold）/ Label fire trigger, width tTriggerHold
    uLabelsApplied : UDINT;                       // 已出标计数 [张]，饱和 / Labels applied [pcs], saturating
    bMissedLabel   : BOOL;                        // 漏标标志，锁存至 bReset / Missed-label flag, latched until reset
    fPhaseErrMm    : LREAL;                       // 相位误差 [mm]，相对出标点：负 = 尚差，正 = 已滞后 / Phase error [mm] relative to the fire point
    fWebSpeedMpm   : LREAL;                       // 卷材线速度 [米每分] / Web line speed [m per min]
    bLowSpeed      : BOOL;                        // 低速抑制出标标志 / Low-speed firing suppression flag
    eErr           : UDINT;                       // 错误码，0 = 无错，码位 16#0004_01ED 起信息级、16#0004_030F 起故障级（分带见错误码表） / Error code, 0 = no error, band info/fault per the code table
    bError         : BOOL;                        // 故障级标志，仅故障级错误置位 / Fault-class flag, set only on fault-level codes
    bValid         : BOOL;                        // 出标扳机可用标志，失能/故障闸显式 FALSE / Trigger usable flag, explicit FALSE on disable/fault gates
    eState         : E_DL_LabelSyncState;         // 主状态机当前状态 / Current state of the main state machine
END_VAR
VAR
    fbReset        : R_TRIG;                      // 复位上升沿检测实例 / Reset rising edge detector
    fbTonHold      : TON;                         // 触发脉宽定时器实例 / Trigger pulse width timer
    nPrevPulse     : DINT;                        // 上拍累计脉冲 [脉冲] / Previous accumulated pulses [pulse]
    nDeltaPulse    : DINT;                        // 本拍脉冲差分 [脉冲]，带符号 / Pulse delta of this scan [pulse], signed
    fDeltaMm       : LREAL;                       // 本拍位移 [mm]，带符号 / Displacement of this scan [mm], signed
    fPhaseMm       : LREAL;                       // 距上次出标的累计相位 [mm] / Accumulated phase since the last fire [mm]
    fTrigPointMm   : LREAL;                       // 出标相位点 = 节距 − 生效提前量 [mm] / Fire phase point [mm]
    fLeadEff       : LREAL;                       // 生效提前量（钳位后）[mm] / Effective lead after clamping [mm]
    fDtSec         : LREAL;                       // 扫描间隔换算成秒 [s] / Scan interval in seconds [s]
    fAbsDeltaMm    : LREAL;                       // 位移绝对值 [mm]，算线速度用 / Absolute displacement for the speed [mm]
    uDtEff         : UDINT;                       // 钳位后的扫描间隔 [ms] / Clamped scan interval [ms]
    bTrigReq       : BOOL;                        // 出标请求（脉宽未撤前后保持）/ Fire request held until the pulse width elapses
    bLeadClamped   : BOOL;                        // 提前量饱和钳位标志 / Lead saturation flag
    bFirstScan     : BOOL := TRUE;                // 上电首拍标志 / First-scan flag
END_VAR
VAR CONSTANT
    DL_LAS_CODE_INFO_1 : UDINT := 16#0004_01ED;   // 信息级槽 1（提前量饱和钳位） / info slot 1
    DL_LAS_CODE_INFO_2 : UDINT := 16#0004_01EE;   // 信息级槽 2（编码器低速暂停出标） / info slot 2
    DL_LAS_CODE_FLT_1  : UDINT := 16#0004_030F;   // 故障级槽 1（脉冲当量/节距组态非法） / fault slot 1
    DL_LAS_CODE_FLT_2  : UDINT := 16#0004_0310;   // 故障级槽 2（输入非有限） / fault slot 2
    DL_LAS_CODE_FLT_3  : UDINT := 16#0004_0311;   // 故障级槽 3（非法状态兜底） / fault slot 3, illegal-state fallback
    DL_LAS_CNT_MAX     : UDINT := 16#FFFF_FFFE;   // 出标计数饱和值 [张] / Label counter saturation [pcs]
    DL_LAS_DT_MIN_MS   : UDINT := 1;              // 扫描间隔下限 [ms]，防除零与死判 / Scan interval floor [ms], prevents divide-by-zero
    DL_LAS_MS_PER_S    : LREAL := 1000.0;         // 毫秒转秒系数 [ms/s] / Milliseconds per second
    DL_LAS_MM_PER_M    : LREAL := 1000.0;         // 毫米转米系数 [mm/m] / Millimetres per metre
    DL_LAS_S_PER_MIN   : LREAL := 60.0;           // 秒转分系数 [s/min] / Seconds per minute
    DL_LAS_ZERO        : LREAL := 0.0;            // 零值常量，避免裸字面量 [—] / Zero constant, avoids a bare literal
    DL_LAS_TOL         : LREAL := 1.0E-6;         // 浮点比较容差 [—] / Float comparison tolerance
    DL_LAS_INF         : LREAL := 1.7976931348623157E308; // LREAL 幅值上限，Inf 判据 / LREAL magnitude ceiling
END_VAR

(*------------------------------------------------------------------------------
 * 段 1｜无条件刷新区（红线 5）：复位沿与脉宽定时器在任何分支之外周期调用
 *----------------------------------------------------------------------------*)
fbReset(CLK := bReset);                            // 复位沿检测无条件刷新 / reset edge refreshed unconditionally
fbTonHold(IN := bTrigReq, PT := tTriggerHold);     // 脉宽定时器无条件刷新 / pulse-width timer refreshed unconditionally

(*------------------------------------------------------------------------------
 * 段 2｜复位沿处理（改写置于沿后，防吞沿 R39）：清漏标锁存与计数并重新对齐相位
 *----------------------------------------------------------------------------*)
IF fbReset.Q THEN
    eState := E_DL_LabelSyncState.eIdle;
    eErr   := 16#0000_0000;                        // 复位清码 / reset clears the code
    bError := FALSE;                               // 复位清故障 / reset clears the fault
    bMissedLabel := FALSE;                         // 漏标锁存清 / missed-label latch cleared
    bLeadClamped := FALSE;                         // 饱和提示清 / saturation hint cleared
    uLabelsApplied := 16#0000_0000;                // 出标计数清 / label counter cleared
    fPhaseMm := DL_LAS_ZERO;                       // 相位清零 / phase cleared
    bTrigReq := FALSE;                             // 出标请求清 / fire request cleared
    bFirstScan := TRUE;                            // 重新首拍化（相位基准重新对齐）/ re-initialize first scan, phase re-based
END_IF

(*------------------------------------------------------------------------------
 * 段 3｜非有限输入闸（NaN 自反判 + Inf 幅值上限判，R79）
 *----------------------------------------------------------------------------*)
IF (fPulsePerMm <> fPulsePerMm) OR (ABS(fPulsePerMm) >= DL_LAS_INF)
   OR (fLabelPitchMm <> fLabelPitchMm) OR (ABS(fLabelPitchMm) >= DL_LAS_INF)
   OR (fLeadMm <> fLeadMm) OR (ABS(fLeadMm) >= DL_LAS_INF)
   OR (fSpeedMinMpm <> fSpeedMinMpm) OR (ABS(fSpeedMinMpm) >= DL_LAS_INF) THEN
    eState := E_DL_LabelSyncState.eFault;          // 进故障相 / enter fault state
    eErr   := DL_LAS_CODE_FLT_2;                   // 故障级：输入非有限 / fault: non-finite input
    bError := TRUE;                                // 故障级必置 bError（R45 配对）/ fault-class pairs with bError
    bValid := FALSE;                               // 扳机不可用 / trigger unusable
    bFireTrigger := FALSE;                         // 扳机撤安全侧 / trigger dropped, safe side
    bTrigReq := FALSE;                             // 请求撤 / request dropped
    bLowSpeed := FALSE;                            // 低速标志撤 / low-speed flag withdrawn
    fPhaseErrMm := DL_LAS_ZERO;                    // 相位误差回零 / phase error zeroed
    fWebSpeedMpm := DL_LAS_ZERO;                   // 线速度回零 / web speed zeroed
    RETURN;
END_IF

(*------------------------------------------------------------------------------
 * 段 4｜组态合法性闸：脉冲当量与节距必须为正——本件全部除法严格位于此闸之后
 *       （先判后除，禁把判零写在除子表达式里）
 *----------------------------------------------------------------------------*)
IF (fPulsePerMm <= DL_LAS_TOL) OR (fLabelPitchMm <= DL_LAS_TOL) THEN
    eState := E_DL_LabelSyncState.eFault;          // 进故障相 / enter fault state
    eErr   := DL_LAS_CODE_FLT_1;                   // 故障级：脉冲当量/节距组态非法 / fault: pulse equivalent or pitch invalid
    bError := TRUE;                                // 故障级必置 bError（R45 配对）/ fault-class pairs with bError
    bValid := FALSE;                               // 扳机不可用 / trigger unusable
    bFireTrigger := FALSE;                         // 扳机撤安全侧 / trigger dropped, safe side
    bTrigReq := FALSE;                             // 请求撤 / request dropped
    bLowSpeed := FALSE;                            // 低速标志撤 / low-speed flag withdrawn
    fPhaseErrMm := DL_LAS_ZERO;                    // 相位误差回零 / phase error zeroed
    fWebSpeedMpm := DL_LAS_ZERO;                   // 线速度回零 / web speed zeroed
    RETURN;
END_IF

(*------------------------------------------------------------------------------
 * 段 5｜提前量饱和钳位：提前量不得超一个节距（超出会让出标点跑到上一节距之前）
 *----------------------------------------------------------------------------*)
fLeadEff := fLeadMm;                               // 先取引脚值 / take the pin value first
bLeadClamped := FALSE;                             // 饱和标志逐拍重判 / saturation flag re-judged per scan
IF fLeadEff > fLabelPitchMm - DL_LAS_TOL THEN
    fLeadEff := fLabelPitchMm;                     // 钳到节距（出标点落在相位 0）/ clamped to one pitch, fire point at phase zero
    bLeadClamped := TRUE;                          // 饱和标志置位 / saturation flag raised
END_IF
IF fLeadEff < DL_LAS_ZERO THEN
    fLeadEff := DL_LAS_ZERO;                       // 负提前量钳到零（不提前即到位出标）/ negative lead clamped to zero
    bLeadClamped := TRUE;                          // 越界同样提示 / out-of-range hint raised
END_IF
fTrigPointMm := fLabelPitchMm - fLeadEff;          // 出标相位点 [mm] / fire phase point [mm]

(*------------------------------------------------------------------------------
 * 段 6｜脉冲差分与线速度：nDelta := nNow − nPrev，DINT 回绕时补码减法自然正确，
 *       禁止用 ABS(nNow − nPrev) 之类绝对值比较（正反转会被抹平）
 *----------------------------------------------------------------------------*)
IF bFirstScan THEN
    nPrevPulse := nEncoderPulse;                   // 上电首拍以当前脉冲为基准 / first scan re-bases on the current pulse
    bFirstScan := FALSE;                           // 首拍标志清除 / first-scan flag cleared
END_IF
nDeltaPulse := nEncoderPulse - nPrevPulse;         // 本拍脉冲差分（带符号，回绕安全）[脉冲] / signed pulse delta, wrap safe
nPrevPulse := nEncoderPulse;                       // 基准刷新 / refresh the reference
fDeltaMm := DINT_TO_LREAL(nDeltaPulse) / fPulsePerMm;   // 位移（除子已由段 4 保证为正）[mm] / displacement, divisor proven positive
IF uDeltaTimeMs < DL_LAS_DT_MIN_MS THEN
    uDtEff := DL_LAS_DT_MIN_MS;                    // 间隔过小按 1 ms 下限 / floored interval
ELSE
    uDtEff := uDeltaTimeMs;                        // 间隔原值 / interval as-is
END_IF
fDtSec := UDINT_TO_LREAL(uDtEff) / DL_LAS_MS_PER_S;    // 间隔换算成秒 [s] / interval in seconds
fAbsDeltaMm := ABS(fDeltaMm);                      // 位移绝对值 [mm] / absolute displacement
IF fDtSec > DL_LAS_TOL THEN
    fWebSpeedMpm := fAbsDeltaMm / fDtSec / DL_LAS_MM_PER_M * DL_LAS_S_PER_MIN;   // 线速度 [米每分] / web speed [m per min]
ELSE
    fWebSpeedMpm := DL_LAS_ZERO;                   // 间隔不可用时线速度记零 / speed reads zero when the interval is unusable
END_IF
IF (fWebSpeedMpm <> fWebSpeedMpm) OR (ABS(fWebSpeedMpm) >= DL_LAS_INF) THEN
    fWebSpeedMpm := DL_LAS_ZERO;                   // 解算非有限兜到零（诊断量不冒充有效值）/ non-finite falls back to zero
END_IF

(*------------------------------------------------------------------------------
 * 段 7｜相位累计与出标判据：低速时只累计不出标（回速后按相位补出，不丢位置）；
 *       每拍最多出一次标，残余相位留待下一拍（不写 WHILE，避免单拍突发多标）
 *----------------------------------------------------------------------------*)
IF bEnable THEN
    fPhaseMm := fPhaseMm + fDeltaMm;               // 相位累计（正反转自然增减）[mm] / phase accumulation, signed
END_IF
bLowSpeed := (fWebSpeedMpm < fSpeedMinMpm);        // 低速判据 [米每分] / low-speed predicate [m per min]
IF bTrigReq AND fbTonHold.Q THEN
    bTrigReq := FALSE;                             // 脉宽到点撤请求（单拍标志自清）/ request cleared when the pulse width elapses
END_IF
IF bEnable AND (NOT bLowSpeed) AND bLabelPresent AND (NOT bTrigReq)
   AND (fPhaseMm >= fTrigPointMm - DL_LAS_TOL) THEN
    bTrigReq := TRUE;                              // 出标请求置位（脉宽由定时器收口）/ fire request raised, width bounded by the timer
    fPhaseMm := fPhaseMm - fLabelPitchMm;          // 相位扣一个节距，残余留待下一拍补出 / phase reduced by one pitch, the residual fires later
    IF uLabelsApplied < DL_LAS_CNT_MAX THEN
        uLabelsApplied := uLabelsApplied + 1;      // 出标计数饱和自增 [张] / saturating label increment
    END_IF
END_IF
IF bEnable AND (NOT bLabelPresent) THEN
    bMissedLabel := TRUE;                          // 缺标锁存（本拍不出标，等补标）/ missing-label latched, no fire
END_IF
IF fPhaseMm > fLabelPitchMm THEN
    fPhaseMm := fPhaseMm - fLabelPitchMm;          // 相位越一个节距仍未出标：钳回一节距内，防累计漂移 / one-pitch guard against unbounded phase drift
    bMissedLabel := TRUE;                          // 越节距即漏标 / overrunning a pitch is a missed label
END_IF
fPhaseErrMm := fPhaseMm - fTrigPointMm;            // 相位误差 [mm]：负 = 尚差，正 = 已过出标点 / phase error, negative = short, positive = past the fire point
bFireTrigger := bTrigReq;                          // 扳机输出（脉宽由定时器收口）/ trigger output, width bounded by the timer

(*------------------------------------------------------------------------------
 * 段 8｜状态机：CASE 含 ELSE 兜底（非法状态 → 0311 + 扳机与许可全撤）
 *----------------------------------------------------------------------------*)
CASE eState OF

    E_DL_LabelSyncState.eIdle:
        bFireTrigger := FALSE;                     // 待机扳机撤 / trigger dropped in idle
        bTrigReq := FALSE;                         // 请求撤 / request dropped
        bValid := FALSE;                           // 失能闸显式不可用（R72）/ explicit FALSE on the disable gate
        bLowSpeed := FALSE;                        // 待机不报低速 / no low-speed hint in idle
        fPhaseErrMm := DL_LAS_ZERO;                // 相位误差回零 / phase error zeroed
        eErr := 16#0000_0000;                      // 待机无错 / no error in idle
        bError := FALSE;                           // 待机无故障 / no fault in idle
        IF bEnable THEN
            fPhaseMm := fTrigPointMm - fLabelPitchMm;   // 重新对齐相位基准（下次到点即出标）/ phase re-based
            eState := E_DL_LabelSyncState.eSync;   // 使能进同步相 / enable enters synchronised firing
        END_IF

    E_DL_LabelSyncState.eSync:
        bValid := TRUE;                            // 扳机可用 / trigger usable
        bError := FALSE;                           // 同步相无故障 / no fault in the synchronised state
        eErr := 16#0000_0000;                      // 同步相先清码 / clear the code first
        IF bLeadClamped THEN
            eErr := DL_LAS_CODE_INFO_1;            // 信息级：提前量饱和钳位 / info: lead saturated
        END_IF
        IF bLowSpeed THEN
            eErr := DL_LAS_CODE_INFO_2;            // 信息级：低速暂停出标（优先于钳位提示）/ info: low speed outranks the lead hint
            eState := E_DL_LabelSyncState.eLowSpeed;   // 转低速抑制相 / enter the low-speed state
        END_IF
        IF NOT bEnable THEN
            eState := E_DL_LabelSyncState.eIdle;   // 失能回待机 / disable returns to idle
            bValid := FALSE;                       // 失能闸显式不可用 / explicit FALSE on the disable gate
            bFireTrigger := FALSE;                 // 扳机撤 / trigger dropped
        END_IF

    E_DL_LabelSyncState.eLowSpeed:
        bValid := FALSE;                           // 低速不出标，扳机不可用（R72）/ no fire at low speed, explicit FALSE
        bFireTrigger := FALSE;                     // 扳机撤（硬出标会贴歪）/ trigger dropped, firing would misplace the label
        bTrigReq := FALSE;                         // 请求撤 / request dropped
        bError := FALSE;                           // 信息级不置 bError（R45/R101）/ info never raises bError
        eErr := DL_LAS_CODE_INFO_2;                // 信息级：编码器低速，无法同步 / info: low speed, cannot synchronise
        IF NOT bEnable THEN
            eState := E_DL_LabelSyncState.eIdle;   // 失能回待机（退出条件一）/ disable, first exit
            bValid := FALSE;                       // 失能闸显式不可用 / explicit FALSE on the disable gate
        ELSIF (NOT bLowSpeed) THEN
            eState := E_DL_LabelSyncState.eSync;   // 速度恢复回同步相（退出条件二）/ speed recovered, second exit
        END_IF

    E_DL_LabelSyncState.eFault:
        bValid := FALSE;                           // 故障闸显式不可用（R72）/ explicit FALSE on the fault gate
        bFireTrigger := FALSE;                     // 扳机撤安全侧 / trigger dropped, safe side
        bTrigReq := FALSE;                         // 请求撤 / request dropped
        bError := TRUE;                            // 故障级必置 bError（R45 配对）/ fault-class pairs with bError
        IF eErr = 16#0000_0000 THEN
            eErr := DL_LAS_CODE_FLT_3;             // 入口无码时按非法状态兜底（R45：bError 必须有对应码）/ illegal-state fallback
        END_IF
        IF bEnable AND (fPulsePerMm > DL_LAS_TOL) AND (fLabelPitchMm > DL_LAS_TOL) THEN
            eState := E_DL_LabelSyncState.eIdle;   // 组态恢复且使能才回待机（退出条件 ≥2）/ recover only when the configuration is sane again
        END_IF

    ELSE
        eState := E_DL_LabelSyncState.eFault;      // 非法状态兜底 / illegal-state fallback
        eErr := DL_LAS_CODE_FLT_3;                 // 故障级兜底：非法状态 / fault fallback: illegal state
        bError := TRUE;                            // 故障级必置 bError（R45 配对）/ fault-class pairs with bError
        bValid := FALSE;                           // 扳机不可用 / trigger unusable
        bFireTrigger := FALSE;                     // 扳机撤安全侧 / trigger dropped, safe side
        bTrigReq := FALSE;                         // 请求撤 / request dropped
        fPhaseErrMm := DL_LAS_ZERO;                // 相位误差回零 / phase error zeroed

END_CASE
END_FUNCTION_BLOCK

(* ---- FB_DL_LamStepperFeed.st ---- *)
// =====================================================================
// FB_DL_LamStepperFeed.st
// 层压机铺膜步进送料（开环步进契约消费 + 膜长累计 + 保养窗冻结 + 堵转判据）
// Laminator film stepper feeding with maintenance freeze and stall judge
// 所属子库: DL_Motion    版本: v1.0.0    兼容: CODESYS V3.5+ / TwinCAT 3 / 汇川 InoProShop
// 码位: 16#0004_0359 ~ 16#0004_035D (本件独占 5 槽, 勿复用)
// 溯源: 道莅 clean-room 防御性实现
//       来源组标签: photovoltaic, laminator, stepper-open-loop, maintenance
// 修改记录: R30 初版 (ROUND_PLAN_R30 序 15)
// 分层声明: 本件为组合编排件, 开环步进运动语义全部经引脚注入消费
//           （就绪/完成/故障回读对应开环步进契约, 不自造轴状态枚举）;
//           累计送料经定长计米件注入; 保养窗经保养窗管理件注入
// =====================================================================
FUNCTION_BLOCK FB_DL_LamStepperFeed
VAR_INPUT
    bStepperReady    : BOOL := FALSE;   // 步进驱动就绪回读注入 / Stepper ready feedback injected
    bStepperDone     : BOOL := FALSE;   // 步进完成回读注入 / Stepper done feedback injected
    bStepperFault    : BOOL := FALSE;   // 步进故障回读注入 / Stepper fault feedback injected
    bFeedStart       : BOOL := FALSE;   // 送料步启动命令 / Feed step start command
    fFilmLen_m       : REAL := 300.0;   // 单卷膜长 0~2000 m / Film roll length [m]
    fStepLen_m       : REAL := 0.5;     // 单步步长 0~10 m / Step length [m]
    fChangeReserve_m : REAL := 5.0;     // 换膜余量 0~50 m / Change reserve [m]
    fFedLen_m        : REAL := 0.0;     // 累计送料反馈注入 0~2000 m / Fed length feedback injected [m]
    bMaintWin        : BOOL := FALSE;   // 保养窗激活注入 / Maintenance window injected
    tFeedTimeout     : TIME := T#10S;   // 送料超时窗（理论耗时×1.5 口径）T#100MS~T#120S / Feed timeout [s]
END_VAR
VAR_OUTPUT
    bFeedCmd    : BOOL := FALSE;        // 送料指令输出 / Feed command output
    bFeedDone   : BOOL := FALSE;        // 步完成脉冲（单拍自清）/ Step done pulse, one cycle
    fRemainLen_m: REAL := 0.0;          // 剩余膜长 / Remaining film length [m]
    bMaintHold  : BOOL := FALSE;        // 保养窗冻结标志（安全侧不启动）/ Maintenance hold flag
    eErr        : UDINT := 16#0004_0359;  // 错误码 / Error code
END_VAR
VAR
    rtrStart  : R_TRIG;                 // 启动沿检测, 每拍无条件刷新 / Start edge, refreshed every cycle
    rtrDone   : R_TRIG;                 // 完成沿检测, 每拍无条件刷新 / Done edge, refreshed every cycle
    tonFeed   : TON;                    // 送料超时定时器, 每拍无条件刷新 / Feed timeout timer, refreshed every cycle
    xFeedAct  : BOOL := FALSE;          // 送料步进行中标志 / Feed step active flag
    bTmoLatch : BOOL := FALSE;          // 超时堵转锁存 / Timeout stall latch
    bCfgErr   : BOOL := FALSE;          // 组态非法标记 / Configuration error flag
    bWarn     : BOOL := FALSE;          // 膜长耗尽预警标记 / Film-end warning flag
END_VAR

// ---------------------------------------------------------------------
// 代码位表（本件独占, 勿复用）:
//   16#0004_0359 信息 送料正常
//   16#0004_035A 故障 送料超时判堵转（指令后未在窗内完成, 指令立即收口）,
//                解除式 = 步进就绪恢复 且 送料步已收口
//   16#0004_035B 故障 步进驱动故障回读有效（指令立即收口）,
//                解除式 = 故障回读消失
//   16#0004_035C 信息 膜长耗尽预警（剩余膜长低于换膜余量, 送料继续）
//   16#0004_035D 故障 组态非法（膜长/步长/余量非有限或不大于 0）,
//                解除式 = 恢复合法组态
// ---------------------------------------------------------------------

// ---- 边沿与定时器实例无条件周期刷新 / Unconditional edge and timer refresh ----
rtrStart(CLK := bFeedStart);        // 启动沿 / Start edge
rtrDone(CLK := bStepperDone);       // 完成沿 / Done edge
tonFeed(IN := xFeedAct, PT := tFeedTimeout);    // 超时计时 / Timeout timing

// ---- 组态闸 / Configuration gate ----
bCfgErr := FALSE;
IF (fFilmLen_m <> fFilmLen_m) OR (fFilmLen_m <= 0.0) OR (fFilmLen_m > 2000.0) THEN
    bCfgErr := TRUE;                // 膜长非法 / Illegal film length
END_IF
IF (fStepLen_m <> fStepLen_m) OR (fStepLen_m <= 0.0) OR (fStepLen_m > 10.0) THEN
    bCfgErr := TRUE;                // 步长非法 / Illegal step length
END_IF
IF (fChangeReserve_m <> fChangeReserve_m) OR (fChangeReserve_m <= 0.0) OR (fChangeReserve_m > 50.0) THEN
    bCfgErr := TRUE;                // 余量非法 / Illegal reserve
END_IF
IF (fFedLen_m <> fFedLen_m) OR (fFedLen_m < 0.0) THEN
    bCfgErr := TRUE;                // 累计送料非法 / Illegal fed length
END_IF

// ---- 保养窗冻结（安全侧: 冻结期指令保持断开）/ Maintenance freeze, safe side ----
bMaintHold := bMaintWin;

// ---- 剩余膜长（负差钳零）/ Remaining film length, negative clamped ----
fRemainLen_m := fFilmLen_m - fFedLen_m;
IF fRemainLen_m < 0.0 THEN
    fRemainLen_m := 0.0;            // 负差钳零 / Clamp to zero
END_IF

// ---- 超时堵转锁存与解除 / Timeout stall latch and release ----
IF tonFeed.Q THEN
    bTmoLatch := TRUE;              // 窗内未完成判堵转锁存 / Stall latch
END_IF
IF bStepperReady AND (NOT xFeedAct) THEN
    bTmoLatch := FALSE;             // 就绪恢复且步已收口 → 解除 / Release on ready recovery
END_IF

// ---- 输出缺省（完成脉冲单拍自清）/ Output defaults, done pulse self-clearing ----
bFeedCmd  := FALSE;
bFeedDone := FALSE;

// ---- 启动沿派步（保养冻结/组态错/堵转/驱动故障/膜尽均不派）/ Start dispatch ----
IF rtrStart.Q AND (NOT bMaintHold) AND (NOT bCfgErr) AND (NOT bTmoLatch)
   AND (NOT bStepperFault) AND bStepperReady AND (fRemainLen_m > 0.0) AND (NOT xFeedAct) THEN
    xFeedAct := TRUE;               // 拍 N 进入送料步 / Enter feed step
END_IF

// ---- 送料步执行与收口 / Feed step execution and closing ----
IF xFeedAct THEN
    IF bMaintHold OR bCfgErr OR bStepperFault THEN
        xFeedAct := FALSE;          // 冻结或故障立即收口（安全侧指令断）/ Close on freeze or fault
    ELSE
        bFeedCmd := TRUE;           // 指令输出 / Command on
        IF rtrDone.Q THEN
            bFeedDone := TRUE;      // 单拍完成脉冲 / One-cycle done pulse
            xFeedAct := FALSE;      // 拍 N+1 步收口 / Close step
        ELSIF tonFeed.Q THEN
            xFeedAct := FALSE;      // 超时收口, 锁存已置 / Close on timeout
        END_IF
    END_IF
END_IF

// ---- 膜长耗尽预警（低于换膜余量, 送料继续）/ Film-end warning, feeding continues ----
bWarn := fRemainLen_m < fChangeReserve_m;

// ---- 错误码仲裁 / Error arbitration ----
IF bCfgErr THEN
    eErr := 16#0004_035D;           // 组态非法 / Config fault
ELSIF bTmoLatch THEN
    eErr := 16#0004_035A;           // 堵转锁存回放 / Stall latch replay
ELSIF bStepperFault THEN
    eErr := 16#0004_035B;           // 驱动故障 / Drive fault
ELSIF bWarn THEN
    eErr := 16#0004_035C;           // 耗尽预警 / Film-end warning
ELSE
    eErr := 16#0004_0359;           // 送料正常 / Feeding normal
END_IF

END_FUNCTION_BLOCK
